//-----------------------------------------------------------------------------------------------------------------------------------------
// PRC 03 Cell loading
//-----------------------------------------------------------------------------------------------------------------------------------------
FOR nStationParameter := 20 TO 35
DO
  GVL_XTS.StationParameter[nStationParameter].rVelo               := 1000.0; //MAIN_APP.rDefaultVeloMin;
END_FOR
nStationParameter := 20;
GVL_XTS.StationParameter[nStationParameter].eType                 := E_STATION_TYPE.STATION_PROCESS;
GVL_XTS.StationParameter[nStationParameter].sText                 := 'PROCESS_INFEED_01';
GVL_XTS.StationParameter[nStationParameter].nConfiguredStopCount  :=       1;   // how many stops the mover has to make in this station

GVL_XTS.StationParameter[nStationParameter].rPosWait              :=    10000.0+80.0; // absolute modulo position
GVL_XTS.StationParameter[nStationParameter].rPosStop[1]           :=       0.0; // relative to rPosWait
GVL_XTS.StationParameter[nStationParameter].rReleaseDistance      :=    1120.0; // relative to Mover.ActPos

nStationParameter := 21;
GVL_XTS.StationParameter[nStationParameter].eType                 := E_STATION_TYPE.STATION_PROCESS;
GVL_XTS.StationParameter[nStationParameter].sText                 := 'PROCESS_INFEED_02';
GVL_XTS.StationParameter[nStationParameter].nConfiguredStopCount  :=       1;   // how many stops the mover has to make in this station

GVL_XTS.StationParameter[nStationParameter].rPosWait              :=    10000.0+160.0; // absolute modulo position
GVL_XTS.StationParameter[nStationParameter].rPosStop[1]           :=       0.0; // relative to rPosWait
GVL_XTS.StationParameter[nStationParameter].rReleaseDistance      :=    1040.0; // relative to Mover.ActPos

nStationParameter := 22;
GVL_XTS.StationParameter[nStationParameter].eType                 := E_STATION_TYPE.STATION_PROCESS;
GVL_XTS.StationParameter[nStationParameter].sText                 := 'PROCESS_INFEED_03';
GVL_XTS.StationParameter[nStationParameter].nConfiguredStopCount  :=       1;   // how many stops the mover has to make in this station

GVL_XTS.StationParameter[nStationParameter].rPosWait              :=    10000.0+240.0; // absolute modulo position
GVL_XTS.StationParameter[nStationParameter].rPosStop[1]           :=       0.0; // relative to rPosWait
GVL_XTS.StationParameter[nStationParameter].rReleaseDistance      :=     960.0; // relative to Mover.ActPos

nStationParameter := 23;
GVL_XTS.StationParameter[nStationParameter].eType                 := E_STATION_TYPE.STATION_PROCESS;
GVL_XTS.StationParameter[nStationParameter].sText                 := 'PROCESS_INFEED_04';
GVL_XTS.StationParameter[nStationParameter].nConfiguredStopCount  :=       1;   // how many stops the mover has to make in this station

GVL_XTS.StationParameter[nStationParameter].rPosWait              :=    10000.0+320.0; // absolute modulo position
GVL_XTS.StationParameter[nStationParameter].rPosStop[1]           :=       0.0; // relative to rPosWait
GVL_XTS.StationParameter[nStationParameter].rReleaseDistance      :=     880.0; // relative to Mover.ActPos

nStationParameter := 24;
GVL_XTS.StationParameter[nStationParameter].eType                 := E_STATION_TYPE.STATION_PROCESS;
GVL_XTS.StationParameter[nStationParameter].sText                 := 'PROCESS_INFEED_05';
GVL_XTS.StationParameter[nStationParameter].nConfiguredStopCount  :=       1;   // how many stops the mover has to make in this station

GVL_XTS.StationParameter[nStationParameter].rPosWait              :=    10000.0+400.0; // absolute modulo position
GVL_XTS.StationParameter[nStationParameter].rPosStop[1]           :=       0.0; // relative to rPosWait
GVL_XTS.StationParameter[nStationParameter].rReleaseDistance      :=     800.0; // relative to Mover.ActPos

nStationParameter := 25;
GVL_XTS.StationParameter[nStationParameter].eType                 := E_STATION_TYPE.STATION_PROCESS;
GVL_XTS.StationParameter[nStationParameter].sText                 := 'PROCESS_INFEED_06';
GVL_XTS.StationParameter[nStationParameter].nConfiguredStopCount  :=       1;   // how many stops the mover has to make in this station

GVL_XTS.StationParameter[nStationParameter].rPosWait              :=    10000.0+480.0; // absolute modulo position
GVL_XTS.StationParameter[nStationParameter].rPosStop[1]           :=       0.0; // relative to rPosWait
GVL_XTS.StationParameter[nStationParameter].rReleaseDistance      :=     720.0; // relative to Mover.ActPos

nStationParameter := 26;
GVL_XTS.StationParameter[nStationParameter].eType                 := E_STATION_TYPE.STATION_PROCESS;
GVL_XTS.StationParameter[nStationParameter].sText                 := 'PROCESS_INFEED_07';
GVL_XTS.StationParameter[nStationParameter].nConfiguredStopCount  :=       1;   // how many stops the mover has to make in this station

GVL_XTS.StationParameter[nStationParameter].rPosWait              :=    10000.0+560.0; // absolute modulo position
GVL_XTS.StationParameter[nStationParameter].rPosStop[1]           :=       0.0; // relative to rPosWait
GVL_XTS.StationParameter[nStationParameter].rReleaseDistance      :=     640.0; // relative to Mover.ActPos

nStationParameter := 27;
GVL_XTS.StationParameter[nStationParameter].eType                 := E_STATION_TYPE.STATION_PROCESS;
GVL_XTS.StationParameter[nStationParameter].sText                 := 'PROCESS_INFEED_08';
GVL_XTS.StationParameter[nStationParameter].nConfiguredStopCount  :=       1;   // how many stops the mover has to make in this station

GVL_XTS.StationParameter[nStationParameter].rPosWait              :=    10000.0+640.0; // absolute modulo position
GVL_XTS.StationParameter[nStationParameter].rPosStop[1]           :=       0.0; // relative to rPosWait
GVL_XTS.StationParameter[nStationParameter].rReleaseDistance      :=     560.0; // relative to Mover.ActPos

nStationParameter := 28;
GVL_XTS.StationParameter[nStationParameter].eType                 := E_STATION_TYPE.STATION_PROCESS;
GVL_XTS.StationParameter[nStationParameter].sText                 := 'PROCESS_INFEED_09';
GVL_XTS.StationParameter[nStationParameter].nConfiguredStopCount  :=       1;   // how many stops the mover has to make in this station

GVL_XTS.StationParameter[nStationParameter].rPosWait              :=    10000.0+720.0; // absolute modulo position
GVL_XTS.StationParameter[nStationParameter].rPosStop[1]           :=       0.0; // relative to rPosWait
GVL_XTS.StationParameter[nStationParameter].rReleaseDistance      :=     480.0; // relative to Mover.ActPos

nStationParameter := 29;
GVL_XTS.StationParameter[nStationParameter].eType                 := E_STATION_TYPE.STATION_PROCESS;
GVL_XTS.StationParameter[nStationParameter].sText                 := 'PROCESS_INFEED_10';
GVL_XTS.StationParameter[nStationParameter].nConfiguredStopCount  :=       1;   // how many stops the mover has to make in this station

GVL_XTS.StationParameter[nStationParameter].rPosWait              :=    10000.0+800.0; // absolute modulo position
GVL_XTS.StationParameter[nStationParameter].rPosStop[1]           :=       0.0; // relative to rPosWait
GVL_XTS.StationParameter[nStationParameter].rReleaseDistance      :=     400.0; // relative to Mover.ActPos

nStationParameter := 30;
GVL_XTS.StationParameter[nStationParameter].eType                 := E_STATION_TYPE.STATION_PROCESS;
GVL_XTS.StationParameter[nStationParameter].sText                 := 'PROCESS_INFEED_11';
GVL_XTS.StationParameter[nStationParameter].nConfiguredStopCount  :=       1;   // how many stops the mover has to make in this station

GVL_XTS.StationParameter[nStationParameter].rPosWait              :=    10000.0+880.0; // absolute modulo position
GVL_XTS.StationParameter[nStationParameter].rPosStop[1]           :=       0.0; // relative to rPosWait
GVL_XTS.StationParameter[nStationParameter].rReleaseDistance      :=     320.0; // relative to Mover.ActPos

nStationParameter := 31;
GVL_XTS.StationParameter[nStationParameter].eType                 := E_STATION_TYPE.STATION_PROCESS;
GVL_XTS.StationParameter[nStationParameter].sText                 := 'PROCESS_INFEED_12';
GVL_XTS.StationParameter[nStationParameter].nConfiguredStopCount  :=       1;   // how many stops the mover has to make in this station

GVL_XTS.StationParameter[nStationParameter].rPosWait              :=    10000.0+960.0; // absolute modulo position
GVL_XTS.StationParameter[nStationParameter].rPosStop[1]           :=       0.0; // relative to rPosWait
GVL_XTS.StationParameter[nStationParameter].rReleaseDistance      :=     240.0; // relative to Mover.ActPos

nStationParameter := 32;
GVL_XTS.StationParameter[nStationParameter].eType                 := E_STATION_TYPE.STATION_PROCESS;
GVL_XTS.StationParameter[nStationParameter].sText                 := 'PROCESS_INFEED_13';
GVL_XTS.StationParameter[nStationParameter].nConfiguredStopCount  :=       1;   // how many stops the mover has to make in this station

GVL_XTS.StationParameter[nStationParameter].rPosWait              :=    10000.0+1040.0; // absolute modulo position
GVL_XTS.StationParameter[nStationParameter].rPosStop[1]           :=       0.0; // relative to rPosWait
GVL_XTS.StationParameter[nStationParameter].rReleaseDistance      :=     160.0; // relative to Mover.ActPos

nStationParameter := 33;
GVL_XTS.StationParameter[nStationParameter].eType                 := E_STATION_TYPE.STATION_PROCESS;
GVL_XTS.StationParameter[nStationParameter].sText                 := 'PROCESS_INFEED_14';
GVL_XTS.StationParameter[nStationParameter].nConfiguredStopCount  :=       1;   // how many stops the mover has to make in this station

GVL_XTS.StationParameter[nStationParameter].rPosWait              :=    10000.0+1120.0; // absolute modulo position
GVL_XTS.StationParameter[nStationParameter].rPosStop[1]           :=       0.0; // relative to rPosWait
GVL_XTS.StationParameter[nStationParameter].rReleaseDistance      :=      80.0; // relative to Mover.ActPos

nStationParameter := 34;
GVL_XTS.StationParameter[nStationParameter].eType                 := E_STATION_TYPE.STATION_PROCESS;
GVL_XTS.StationParameter[nStationParameter].sText                 := 'PROCESS_INFEED_15';
GVL_XTS.StationParameter[nStationParameter].nConfiguredStopCount  :=       1;   // how many stops the mover has to make in this station

GVL_XTS.StationParameter[nStationParameter].rPosWait              :=    10000.0+1200.0; // absolute modulo position
GVL_XTS.StationParameter[nStationParameter].rPosStop[1]           :=       0.0; // relative to rPosWait
GVL_XTS.StationParameter[nStationParameter].rReleaseDistance      :=      25.0; // relative to Mover.ActPos

nStationParameter := 35;
GVL_XTS.StationParameter[nStationParameter].eType                 := E_STATION_TYPE.STATION_PROCESS;
GVL_XTS.StationParameter[nStationParameter].sText                 := 'PROCESS_INFEED_16';
GVL_XTS.StationParameter[nStationParameter].nConfiguredStopCount  :=       1;   // how many stops the mover has to make in this station

GVL_XTS.StationParameter[nStationParameter].rPosWait              :=    10000.0+1280.0; // absolute modulo position
GVL_XTS.StationParameter[nStationParameter].rPosStop[1]           :=       0.0; // relative to rPosWait
GVL_XTS.StationParameter[nStationParameter].rReleaseDistance      :=      -5.0; // relative to Mover.ActPos

//-----------------------------------------------------------------------------------------------------------------------------------------
// CONTINUOUS_CLEAN
//-----------------------------------------------------------------------------------------------------------------------------------------
nStationParameter := 37;
GVL_XTS.StationParameter[nStationParameter].eType                 := E_STATION_TYPE.STATION_PROCESS;
GVL_XTS.StationParameter[nStationParameter].sText                 := 'CONTINUOUS_CLEAN';
GVL_XTS.StationParameter[nStationParameter].nConfiguredStopCount  :=       1;   // how many stops the mover has to make in this station

GVL_XTS.StationParameter[nStationParameter].rPosWait              :=   12900.0; // absolute modulo position
GVL_XTS.StationParameter[nStationParameter].rPosStop[1]           :=       0.0; // relative to rPosWait
GVL_XTS.StationParameter[nStationParameter].rReleaseDistance      :=      -5.0; // relative to Mover.ActPos
GVL_XTS.StationParameter[nStationParameter].rVelo                 :=     250.0;
GVL_XTS.StationParameter[nStationParameter].rGap                  :=     110.0;

//-----------------------------------------------------------------------------------------------------------------------------------------
// CONTINUOUS_SCAN
//-----------------------------------------------------------------------------------------------------------------------------------------
nStationParameter := 38;
GVL_XTS.StationParameter[nStationParameter].eType                 := E_STATION_TYPE.STATION_PROCESS;
GVL_XTS.StationParameter[nStationParameter].sText                 := 'CONTINUOUS_SCAN';
GVL_XTS.StationParameter[nStationParameter].nConfiguredStopCount  :=       1;   // how many stops the mover has to make in this station

GVL_XTS.StationParameter[nStationParameter].rPosWait              :=   14000.0; // absolute modulo position
GVL_XTS.StationParameter[nStationParameter].rPosStop[1]           :=       0.0; // relative to rPosWait
GVL_XTS.StationParameter[nStationParameter].rReleaseDistance      :=      -5.0; // relative to Mover.ActPos
GVL_XTS.StationParameter[nStationParameter].rVelo                 :=     250.0;
GVL_XTS.StationParameter[nStationParameter].rGap                  :=     110.0;

//-----------------------------------------------------------------------------------------------------------------------------------------
// CONTINUOUS_CAM
//-----------------------------------------------------------------------------------------------------------------------------------------
nStationParameter := 39;
GVL_XTS.StationParameter[nStationParameter].eType                 := E_STATION_TYPE.STATION_PROCESS;
GVL_XTS.StationParameter[nStationParameter].sText                 := 'CONTINUOUS_CAM';
GVL_XTS.StationParameter[nStationParameter].nConfiguredStopCount  :=       1;   // how many stops the mover has to make in this station

GVL_XTS.StationParameter[nStationParameter].rPosWait              :=   14300.0; // absolute modulo position
GVL_XTS.StationParameter[nStationParameter].rPosStop[1]           :=       0.0; // relative to rPosWait
GVL_XTS.StationParameter[nStationParameter].rReleaseDistance      :=      -5.0; // relative to Mover.ActPos
GVL_XTS.StationParameter[nStationParameter].rVelo                 :=     250.0;
GVL_XTS.StationParameter[nStationParameter].rGap                  :=     109.0;

//-----------------------------------------------------------------------------------------------------------------------------------------
// DISTRIBUTOR_ASSEMBLY_01
//-----------------------------------------------------------------------------------------------------------------------------------------
nStationParameter := 40;
GVL_XTS.StationParameter[nStationParameter].eType                 := E_STATION_TYPE.STATION_PROCESS;
GVL_XTS.StationParameter[nStationParameter].sText                 := 'DISTRIBUTOR_ASSEMBLY_01';
GVL_XTS.StationParameter[nStationParameter].nConfiguredStopCount  :=       1;   // how many stops the mover has to make in this station

GVL_XTS.StationParameter[nStationParameter].rPosWait              :=   15250.0; // absolute modulo position
GVL_XTS.StationParameter[nStationParameter].rPosStop[1]           :=       0.0; // relative to rPosWait
GVL_XTS.StationParameter[nStationParameter].rReleaseDistance      :=      -5.0; // relative to Mover.ActPos
GVL_XTS.StationParameter[nStationParameter].rVelo                 :=    1500.0;
GVL_XTS.StationParameter[nStationParameter].rGap                  :=     109.0;

//-----------------------------------------------------------------------------------------------------------------------------------------
// PRC 05 Visual check film bottom
//-----------------------------------------------------------------------------------------------------------------------------------------
FOR nStationParameter := 41 TO 56
DO
  GVL_XTS.StationParameter[nStationParameter].rVelo               := MAIN_APP.rDefaultVeloMin;
END_FOR
nStationParameter := 41;
GVL_XTS.StationParameter[nStationParameter].eType                 := E_STATION_TYPE.STATION_PROCESS;
GVL_XTS.StationParameter[nStationParameter].sText                 := 'PROCESS_ASSEMBLY_01_01';
GVL_XTS.StationParameter[nStationParameter].nConfiguredStopCount  :=       1;   // how many stops the mover has to make in this station

GVL_XTS.StationParameter[nStationParameter].rPosWait              :=    15500.0+110.0; // absolute modulo position
GVL_XTS.StationParameter[nStationParameter].rPosStop[1]           :=       0.0; // relative to rPosWait
GVL_XTS.StationParameter[nStationParameter].rReleaseDistance      :=    1100.0; // relative to Mover.ActPos
GVL_XTS.StationParameter[nStationParameter].rGap                  :=     109.0;

nStationParameter := 42;
GVL_XTS.StationParameter[nStationParameter].eType                 := E_STATION_TYPE.STATION_PROCESS;
GVL_XTS.StationParameter[nStationParameter].sText                 := 'PROCESS_ASSEMBLY_01_02';
GVL_XTS.StationParameter[nStationParameter].nConfiguredStopCount  :=       1;   // how many stops the mover has to make in this station

GVL_XTS.StationParameter[nStationParameter].rPosWait              :=    15500.0+220.0; // absolute modulo position
GVL_XTS.StationParameter[nStationParameter].rPosStop[1]           :=       0.0; // relative to rPosWait
GVL_XTS.StationParameter[nStationParameter].rReleaseDistance      :=     990.0; // relative to Mover.ActPos
GVL_XTS.StationParameter[nStationParameter].rGap                  :=     109.0;

nStationParameter := 43;
GVL_XTS.StationParameter[nStationParameter].eType                 := E_STATION_TYPE.STATION_PROCESS;
GVL_XTS.StationParameter[nStationParameter].sText                 := 'PROCESS_ASSEMBLY_01_03';
GVL_XTS.StationParameter[nStationParameter].nConfiguredStopCount  :=       1;   // how many stops the mover has to make in this station

GVL_XTS.StationParameter[nStationParameter].rPosWait              :=    15500.0+330.0; // absolute modulo position
GVL_XTS.StationParameter[nStationParameter].rPosStop[1]           :=       0.0; // relative to rPosWait
GVL_XTS.StationParameter[nStationParameter].rReleaseDistance      :=     880.0; // relative to Mover.ActPos
GVL_XTS.StationParameter[nStationParameter].rGap                  :=     109.0;

nStationParameter := 44;
GVL_XTS.StationParameter[nStationParameter].eType                 := E_STATION_TYPE.STATION_PROCESS;
GVL_XTS.StationParameter[nStationParameter].sText                 := 'PROCESS_ASSEMBLY_01_04';
GVL_XTS.StationParameter[nStationParameter].nConfiguredStopCount  :=       1;   // how many stops the mover has to make in this station

GVL_XTS.StationParameter[nStationParameter].rPosWait              :=    15500.0+440.0; // absolute modulo position
GVL_XTS.StationParameter[nStationParameter].rPosStop[1]           :=       0.0; // relative to rPosWait
GVL_XTS.StationParameter[nStationParameter].rReleaseDistance      :=     770.0; // relative to Mover.ActPos
GVL_XTS.StationParameter[nStationParameter].rGap                  :=     109.0;

nStationParameter := 45;
GVL_XTS.StationParameter[nStationParameter].eType                 := E_STATION_TYPE.STATION_PROCESS;
GVL_XTS.StationParameter[nStationParameter].sText                 := 'PROCESS_ASSEMBLY_01_05';
GVL_XTS.StationParameter[nStationParameter].nConfiguredStopCount  :=       1;   // how many stops the mover has to make in this station

GVL_XTS.StationParameter[nStationParameter].rPosWait              :=    15500.0+550.0; // absolute modulo position
GVL_XTS.StationParameter[nStationParameter].rPosStop[1]           :=       0.0; // relative to rPosWait
GVL_XTS.StationParameter[nStationParameter].rReleaseDistance      :=     660.0; // relative to Mover.ActPos
GVL_XTS.StationParameter[nStationParameter].rGap                  :=     109.0;

nStationParameter := 46;
GVL_XTS.StationParameter[nStationParameter].eType                 := E_STATION_TYPE.STATION_PROCESS;
GVL_XTS.StationParameter[nStationParameter].sText                 := 'PROCESS_ASSEMBLY_01_06';
GVL_XTS.StationParameter[nStationParameter].nConfiguredStopCount  :=       1;   // how many stops the mover has to make in this station

GVL_XTS.StationParameter[nStationParameter].rPosWait              :=    15500.0+660.0; // absolute modulo position
GVL_XTS.StationParameter[nStationParameter].rPosStop[1]           :=       0.0; // relative to rPosWait
GVL_XTS.StationParameter[nStationParameter].rReleaseDistance      :=     550.0; // relative to Mover.ActPos
GVL_XTS.StationParameter[nStationParameter].rGap                  :=     109.0;

nStationParameter := 47;
GVL_XTS.StationParameter[nStationParameter].eType                 := E_STATION_TYPE.STATION_PROCESS;
GVL_XTS.StationParameter[nStationParameter].sText                 := 'PROCESS_ASSEMBLY_01_07';
GVL_XTS.StationParameter[nStationParameter].nConfiguredStopCount  :=       1;   // how many stops the mover has to make in this station

GVL_XTS.StationParameter[nStationParameter].rPosWait              :=    15500.0+770.0; // absolute modulo position
GVL_XTS.StationParameter[nStationParameter].rPosStop[1]           :=       0.0; // relative to rPosWait
GVL_XTS.StationParameter[nStationParameter].rReleaseDistance      :=     440.0; // relative to Mover.ActPos
GVL_XTS.StationParameter[nStationParameter].rGap                  :=     109.0;

nStationParameter := 48;
GVL_XTS.StationParameter[nStationParameter].eType                 := E_STATION_TYPE.STATION_PROCESS;
GVL_XTS.StationParameter[nStationParameter].sText                 := 'PROCESS_ASSEMBLY_01_08';
GVL_XTS.StationParameter[nStationParameter].nConfiguredStopCount  :=       1;   // how many stops the mover has to make in this station

GVL_XTS.StationParameter[nStationParameter].rPosWait              :=    15500.0+880.0; // absolute modulo position
GVL_XTS.StationParameter[nStationParameter].rPosStop[1]           :=       0.0; // relative to rPosWait
GVL_XTS.StationParameter[nStationParameter].rReleaseDistance      :=     330.0; // relative to Mover.ActPos
GVL_XTS.StationParameter[nStationParameter].rGap                  :=     109.0;

nStationParameter := 49;
GVL_XTS.StationParameter[nStationParameter].eType                 := E_STATION_TYPE.STATION_PROCESS;
GVL_XTS.StationParameter[nStationParameter].sText                 := 'PROCESS_ASSEMBLY_01_09';
GVL_XTS.StationParameter[nStationParameter].nConfiguredStopCount  :=       1;   // how many stops the mover has to make in this station

GVL_XTS.StationParameter[nStationParameter].rPosWait              :=    15500.0+990.0; // absolute modulo position
GVL_XTS.StationParameter[nStationParameter].rPosStop[1]           :=       0.0; // relative to rPosWait
GVL_XTS.StationParameter[nStationParameter].rReleaseDistance      :=     220.0; // relative to Mover.ActPos
GVL_XTS.StationParameter[nStationParameter].rGap                  :=     109.0;

nStationParameter := 50;
GVL_XTS.StationParameter[nStationParameter].eType                 := E_STATION_TYPE.STATION_PROCESS;
GVL_XTS.StationParameter[nStationParameter].sText                 := 'PROCESS_ASSEMBLY_01_10';
GVL_XTS.StationParameter[nStationParameter].nConfiguredStopCount  :=       1;   // how many stops the mover has to make in this station
GVL_XTS.StationParameter[nStationParameter].rGap                  :=     110.0;

GVL_XTS.StationParameter[nStationParameter].rPosWait              :=    15500.0+1100.0; // absolute modulo position
GVL_XTS.StationParameter[nStationParameter].rPosStop[1]           :=       0.0; // relative to rPosWait
GVL_XTS.StationParameter[nStationParameter].rReleaseDistance      :=     110.0; // relative to Mover.ActPos
GVL_XTS.StationParameter[nStationParameter].rGap                  :=     109.0;

nStationParameter := 51;
GVL_XTS.StationParameter[nStationParameter].eType                 := E_STATION_TYPE.STATION_PROCESS;
GVL_XTS.StationParameter[nStationParameter].sText                 := 'PROCESS_ASSEMBLY_01_11';
GVL_XTS.StationParameter[nStationParameter].nConfiguredStopCount  :=       1;   // how many stops the mover has to make in this station

GVL_XTS.StationParameter[nStationParameter].rPosWait              :=    15500.0+1210.0; // absolute modulo position
GVL_XTS.StationParameter[nStationParameter].rPosStop[1]           :=       0.0; // relative to rPosWait
GVL_XTS.StationParameter[nStationParameter].rReleaseDistance      :=     25.0; // relative to Mover.ActPos
GVL_XTS.StationParameter[nStationParameter].rGap                  :=     109.0;

nStationParameter := 52;
GVL_XTS.StationParameter[nStationParameter].eType                 := E_STATION_TYPE.STATION_PROCESS;
GVL_XTS.StationParameter[nStationParameter].sText                 := 'PROCESS_ASSEMBLY_01_12';
GVL_XTS.StationParameter[nStationParameter].nConfiguredStopCount  :=       1;   // how many stops the mover has to make in this station

GVL_XTS.StationParameter[nStationParameter].rPosWait              :=    15500.0+1320.0; // absolute modulo position
GVL_XTS.StationParameter[nStationParameter].rPosStop[1]           :=       0.0; // relative to rPosWait
GVL_XTS.StationParameter[nStationParameter].rReleaseDistance      :=     330.0; // relative to Mover.ActPos
GVL_XTS.StationParameter[nStationParameter].rGap                  :=     109.0;

nStationParameter := 53;
GVL_XTS.StationParameter[nStationParameter].eType                 := E_STATION_TYPE.STATION_PROCESS;
GVL_XTS.StationParameter[nStationParameter].sText                 := 'PROCESS_ASSEMBLY_01_13';
GVL_XTS.StationParameter[nStationParameter].nConfiguredStopCount  :=       1;   // how many stops the mover has to make in this station

GVL_XTS.StationParameter[nStationParameter].rPosWait              :=    15500.0+1430.0; // absolute modulo position
GVL_XTS.StationParameter[nStationParameter].rPosStop[1]           :=       0.0; // relative to rPosWait
GVL_XTS.StationParameter[nStationParameter].rReleaseDistance      :=     220.0; // relative to Mover.ActPos
GVL_XTS.StationParameter[nStationParameter].rGap                  :=     109.0;

nStationParameter := 54;
GVL_XTS.StationParameter[nStationParameter].eType                 := E_STATION_TYPE.STATION_PROCESS;
GVL_XTS.StationParameter[nStationParameter].sText                 := 'PROCESS_ASSEMBLY_01_14';
GVL_XTS.StationParameter[nStationParameter].nConfiguredStopCount  :=       1;   // how many stops the mover has to make in this station

GVL_XTS.StationParameter[nStationParameter].rPosWait              :=    15500.0+1540.0; // absolute modulo position
GVL_XTS.StationParameter[nStationParameter].rPosStop[1]           :=       0.0; // relative to rPosWait
GVL_XTS.StationParameter[nStationParameter].rReleaseDistance      :=     110.0; // relative to Mover.ActPos
GVL_XTS.StationParameter[nStationParameter].rGap                  :=     109.0;

nStationParameter := 55;
GVL_XTS.StationParameter[nStationParameter].eType                 := E_STATION_TYPE.STATION_PROCESS;
GVL_XTS.StationParameter[nStationParameter].sText                 := 'PROCESS_ASSEMBLY_01_15';
GVL_XTS.StationParameter[nStationParameter].nConfiguredStopCount  :=       1;   // how many stops the mover has to make in this station

GVL_XTS.StationParameter[nStationParameter].rPosWait              :=    15500.0+1650.0; // absolute modulo position
GVL_XTS.StationParameter[nStationParameter].rPosStop[1]           :=       0.0; // relative to rPosWait
GVL_XTS.StationParameter[nStationParameter].rReleaseDistance      :=      25.0; // relative to Mover.ActPos
GVL_XTS.StationParameter[nStationParameter].rGap                  :=     109.0;

nStationParameter := 56;
GVL_XTS.StationParameter[nStationParameter].eType                 := E_STATION_TYPE.STATION_PROCESS;
GVL_XTS.StationParameter[nStationParameter].sText                 := 'PROCESS_ASSEMBLY_01_16';
GVL_XTS.StationParameter[nStationParameter].nConfiguredStopCount  :=       1;   // how many stops the mover has to make in this station

GVL_XTS.StationParameter[nStationParameter].rPosWait              :=    15500.0+1740.0; // absolute modulo position
GVL_XTS.StationParameter[nStationParameter].rPosStop[1]           :=       0.0; // relative to rPosWait
GVL_XTS.StationParameter[nStationParameter].rReleaseDistance      :=      -5.0; // relative to Mover.ActPos
GVL_XTS.StationParameter[nStationParameter].rGap                  :=     109.0;
//-----------------------------------------------------------------------------------------------------------------------------------------
// DISTRIBUTOR_ASSEMBLY_02
//-----------------------------------------------------------------------------------------------------------------------------------------
nStationParameter := 57;
GVL_XTS.StationParameter[nStationParameter].eType                 := E_STATION_TYPE.STATION_PROCESS;
GVL_XTS.StationParameter[nStationParameter].sText                 := 'DISTRIBUTOR_ASSEMBLY_02';
GVL_XTS.StationParameter[nStationParameter].nConfiguredStopCount  :=       1;   // how many stops the mover has to make in this station

GVL_XTS.StationParameter[nStationParameter].rPosWait              :=   18000.0; // absolute modulo position
GVL_XTS.StationParameter[nStationParameter].rPosStop[1]           :=       0.0; // relative to rPosWait
GVL_XTS.StationParameter[nStationParameter].rReleaseDistance      :=      -5.0; // relative to Mover.ActPos
GVL_XTS.StationParameter[nStationParameter].rVelo                 := MAIN_APP.rDefaultVeloMin;

//-----------------------------------------------------------------------------------------------------------------------------------------
// PROCESS_ASSEMBLY_02
//-----------------------------------------------------------------------------------------------------------------------------------------
FOR nStationParameter := 58 TO 69
DO
   GVL_XTS.StationParameter[nStationParameter].rVelo               := MAIN_APP.rDefaultVeloMin;
END_FOR
nStationParameter := 58;
GVL_XTS.StationParameter[nStationParameter].eType                 := E_STATION_TYPE.STATION_PROCESS;
GVL_XTS.StationParameter[nStationParameter].sText                 := 'PROCESS_ASSEMBLY_02_01';
GVL_XTS.StationParameter[nStationParameter].nConfiguredStopCount  :=       1;   // how many stops the mover has to make in this station

GVL_XTS.StationParameter[nStationParameter].rPosWait              :=    19500.0+80.0; // absolute modulo position
GVL_XTS.StationParameter[nStationParameter].rPosStop[1]           :=       0.0; // relative to rPosWait
GVL_XTS.StationParameter[nStationParameter].rReleaseDistance      :=     480.0; // relative to Mover.ActPos

nStationParameter := 59;
GVL_XTS.StationParameter[nStationParameter].eType                 := E_STATION_TYPE.STATION_PROCESS;
GVL_XTS.StationParameter[nStationParameter].sText                 := 'PROCESS_ASSEMBLY_02_02';
GVL_XTS.StationParameter[nStationParameter].nConfiguredStopCount  :=       1;   // how many stops the mover has to make in this station

GVL_XTS.StationParameter[nStationParameter].rPosWait              :=    19500.0+160.0; // absolute modulo position
GVL_XTS.StationParameter[nStationParameter].rPosStop[1]           :=       0.0; // relative to rPosWait
GVL_XTS.StationParameter[nStationParameter].rReleaseDistance      :=     400.0; // relative to Mover.ActPos

nStationParameter := 60;
GVL_XTS.StationParameter[nStationParameter].eType                 := E_STATION_TYPE.STATION_PROCESS;
GVL_XTS.StationParameter[nStationParameter].sText                 := 'PROCESS_ASSEMBLY_02_03';
GVL_XTS.StationParameter[nStationParameter].nConfiguredStopCount  :=       1;   // how many stops the mover has to make in this station

GVL_XTS.StationParameter[nStationParameter].rPosWait              :=    19500.0+240.0; // absolute modulo position
GVL_XTS.StationParameter[nStationParameter].rPosStop[1]           :=       0.0; // relative to rPosWait
GVL_XTS.StationParameter[nStationParameter].rReleaseDistance      :=     320.0; // relative to Mover.ActPos

nStationParameter := 61;
GVL_XTS.StationParameter[nStationParameter].eType                 := E_STATION_TYPE.STATION_PROCESS;
GVL_XTS.StationParameter[nStationParameter].sText                 := 'PROCESS_ASSEMBLY_02_04';
GVL_XTS.StationParameter[nStationParameter].nConfiguredStopCount  :=       1;   // how many stops the mover has to make in this station

GVL_XTS.StationParameter[nStationParameter].rPosWait              :=    19500.0+320.0; // absolute modulo position
GVL_XTS.StationParameter[nStationParameter].rPosStop[1]           :=       0.0; // relative to rPosWait
GVL_XTS.StationParameter[nStationParameter].rReleaseDistance      :=     240.0; // relative to Mover.ActPos

nStationParameter := 62;
GVL_XTS.StationParameter[nStationParameter].eType                 := E_STATION_TYPE.STATION_PROCESS;
GVL_XTS.StationParameter[nStationParameter].sText                 := 'PROCESS_ASSEMBLY_02_05';
GVL_XTS.StationParameter[nStationParameter].nConfiguredStopCount  :=       1;   // how many stops the mover has to make in this station

GVL_XTS.StationParameter[nStationParameter].rPosWait              :=    19500.0+400.0; // absolute modulo position
GVL_XTS.StationParameter[nStationParameter].rPosStop[1]           :=       0.0; // relative to rPosWait
GVL_XTS.StationParameter[nStationParameter].rReleaseDistance      :=      160.0; // relative to Mover.ActPos

nStationParameter := 63;
GVL_XTS.StationParameter[nStationParameter].eType                 := E_STATION_TYPE.STATION_PROCESS;
GVL_XTS.StationParameter[nStationParameter].sText                 := 'PROCESS_ASSEMBLY_02_06';
GVL_XTS.StationParameter[nStationParameter].nConfiguredStopCount  :=       1;   // how many stops the mover has to make in this station

GVL_XTS.StationParameter[nStationParameter].rPosWait              :=    19500.0+480.0; // absolute modulo position
GVL_XTS.StationParameter[nStationParameter].rPosStop[1]           :=       0.0; // relative to rPosWait
GVL_XTS.StationParameter[nStationParameter].rReleaseDistance      :=      80.0; // relative to Mover.ActPos

nStationParameter := 64;
GVL_XTS.StationParameter[nStationParameter].eType                 := E_STATION_TYPE.STATION_PROCESS;
GVL_XTS.StationParameter[nStationParameter].sText                 := 'PROCESS_ASSEMBLY_02_07';
GVL_XTS.StationParameter[nStationParameter].nConfiguredStopCount  :=       1;   // how many stops the mover has to make in this station

GVL_XTS.StationParameter[nStationParameter].rPosWait              :=    19500.0+560.0; // absolute modulo position
GVL_XTS.StationParameter[nStationParameter].rPosStop[1]           :=       0.0; // relative to rPosWait
GVL_XTS.StationParameter[nStationParameter].rReleaseDistance      :=      25.0; // relative to Mover.ActPos

nStationParameter := 65;
GVL_XTS.StationParameter[nStationParameter].eType                 := E_STATION_TYPE.STATION_PROCESS;
GVL_XTS.StationParameter[nStationParameter].sText                 := 'PROCESS_ASSEMBLY_02_08';
GVL_XTS.StationParameter[nStationParameter].nConfiguredStopCount  :=       1;   // how many stops the mover has to make in this station

GVL_XTS.StationParameter[nStationParameter].rPosWait              :=    19500.0+640.0; // absolute modulo position
GVL_XTS.StationParameter[nStationParameter].rPosStop[1]           :=       0.0; // relative to rPosWait
GVL_XTS.StationParameter[nStationParameter].rReleaseDistance      :=     -5.0; // relative to Mover.ActPos

nStationParameter := 66;
GVL_XTS.StationParameter[nStationParameter].eType                 := E_STATION_TYPE.STATION_PROCESS;
GVL_XTS.StationParameter[nStationParameter].sText                 := 'PROCESS_ASSEMBLY_02_09';
GVL_XTS.StationParameter[nStationParameter].nConfiguredStopCount  :=       1;   // how many stops the mover has to make in this station

GVL_XTS.StationParameter[nStationParameter].rPosWait              :=    19500.0+720.0; // absolute modulo position
GVL_XTS.StationParameter[nStationParameter].rPosStop[1]           :=       0.0; // relative to rPosWait
GVL_XTS.StationParameter[nStationParameter].rReleaseDistance      :=     240.0; // relative to Mover.ActPos

nStationParameter := 67;
GVL_XTS.StationParameter[nStationParameter].eType                 := E_STATION_TYPE.STATION_PROCESS;
GVL_XTS.StationParameter[nStationParameter].sText                 := 'PROCESS_ASSEMBLY_02_10';
GVL_XTS.StationParameter[nStationParameter].nConfiguredStopCount  :=       1;   // how many stops the mover has to make in this station

GVL_XTS.StationParameter[nStationParameter].rPosWait              :=    19500.0+800.0; // absolute modulo position
GVL_XTS.StationParameter[nStationParameter].rPosStop[1]           :=       0.0; // relative to rPosWait
GVL_XTS.StationParameter[nStationParameter].rReleaseDistance      :=     160.0; // relative to Mover.ActPos

nStationParameter := 68;
GVL_XTS.StationParameter[nStationParameter].eType                 := E_STATION_TYPE.STATION_PROCESS;
GVL_XTS.StationParameter[nStationParameter].sText                 := 'PROCESS_ASSEMBLY_02_11';
GVL_XTS.StationParameter[nStationParameter].nConfiguredStopCount  :=       1;   // how many stops the mover has to make in this station

GVL_XTS.StationParameter[nStationParameter].rPosWait              :=    19500.0+880.0; // absolute modulo position
GVL_XTS.StationParameter[nStationParameter].rPosStop[1]           :=       0.0; // relative to rPosWait
GVL_XTS.StationParameter[nStationParameter].rReleaseDistance      :=      80.0; // relative to Mover.ActPos

nStationParameter := 69;
GVL_XTS.StationParameter[nStationParameter].eType                 := E_STATION_TYPE.STATION_PROCESS;
GVL_XTS.StationParameter[nStationParameter].sText                 := 'PROCESS_ASSEMBLY_02_12';
GVL_XTS.StationParameter[nStationParameter].nConfiguredStopCount  :=       1;   // how many stops the mover has to make in this station

GVL_XTS.StationParameter[nStationParameter].rPosWait              :=    19500.0+960.0; // absolute modulo position
GVL_XTS.StationParameter[nStationParameter].rPosStop[1]           :=       0.0; // relative to rPosWait
GVL_XTS.StationParameter[nStationParameter].rReleaseDistance      :=      25.0; // relative to Mover.ActPos

//-----------------------------------------------------------------------------------------------------------------------------------------
// DISTRIBUTOR_ASSEMBLY_TEST
//-----------------------------------------------------------------------------------------------------------------------------------------
nStationParameter := 70;
GVL_XTS.StationParameter[nStationParameter].eType                 := E_STATION_TYPE.STATION_PROCESS;
GVL_XTS.StationParameter[nStationParameter].sText                 := 'DISTRIBUTOR_ASSEMBLY_TEST';
GVL_XTS.StationParameter[nStationParameter].nConfiguredStopCount  :=       1;   // how many stops the mover has to make in this station

GVL_XTS.StationParameter[nStationParameter].rPosWait              :=   21000.0; // absolute modulo position
GVL_XTS.StationParameter[nStationParameter].rPosStop[1]           :=       0.0; // relative to rPosWait
GVL_XTS.StationParameter[nStationParameter].rReleaseDistance      :=      -5.0; // relative to Mover.ActPos


//-----------------------------------------------------------------------------------------------------------------------------------------
// PROCESS_ASSEMBLY_TEST
//-----------------------------------------------------------------------------------------------------------------------------------------
FOR nStationParameter := 71 TO 86
DO
   GVL_XTS.StationParameter[nStationParameter].rVelo               := 1000.0;//MAIN_APP.rDefaultVeloMin;
END_FOR
nStationParameter := 71;
GVL_XTS.StationParameter[nStationParameter].eType                 := E_STATION_TYPE.STATION_PROCESS;
GVL_XTS.StationParameter[nStationParameter].sText                 := 'PROCESS_ASSEMBLY_TEST_01';
GVL_XTS.StationParameter[nStationParameter].nConfiguredStopCount  :=       1;   // how many stops the mover has to make in this station

GVL_XTS.StationParameter[nStationParameter].rPosWait              :=    21500.0+80.0; // absolute modulo position
GVL_XTS.StationParameter[nStationParameter].rPosStop[1]           :=       0.0; // relative to rPosWait
GVL_XTS.StationParameter[nStationParameter].rReleaseDistance      :=     800.0; // relative to Mover.ActPos

nStationParameter := 72;
GVL_XTS.StationParameter[nStationParameter].eType                 := E_STATION_TYPE.STATION_PROCESS;
GVL_XTS.StationParameter[nStationParameter].sText                 := 'PROCESS_ASSEMBLY_TEST_02';
GVL_XTS.StationParameter[nStationParameter].nConfiguredStopCount  :=       1;   // how many stops the mover has to make in this station

GVL_XTS.StationParameter[nStationParameter].rPosWait              :=    21500.0+160.0; // absolute modulo position
GVL_XTS.StationParameter[nStationParameter].rPosStop[1]           :=       0.0; // relative to rPosWait
GVL_XTS.StationParameter[nStationParameter].rReleaseDistance      :=     720.0; // relative to Mover.ActPos

nStationParameter := 73;
GVL_XTS.StationParameter[nStationParameter].eType                 := E_STATION_TYPE.STATION_PROCESS;
GVL_XTS.StationParameter[nStationParameter].sText                 := 'PROCESS_ASSEMBLY_TEST_03';
GVL_XTS.StationParameter[nStationParameter].nConfiguredStopCount  :=       1;   // how many stops the mover has to make in this station

GVL_XTS.StationParameter[nStationParameter].rPosWait              :=    21500.0+240.0; // absolute modulo position
GVL_XTS.StationParameter[nStationParameter].rPosStop[1]           :=       0.0; // relative to rPosWait
GVL_XTS.StationParameter[nStationParameter].rReleaseDistance      :=    640.0; // relative to Mover.ActPos

nStationParameter := 74;
GVL_XTS.StationParameter[nStationParameter].eType                 := E_STATION_TYPE.STATION_PROCESS;
GVL_XTS.StationParameter[nStationParameter].sText                 := 'PROCESS_ASSEMBLY_TEST_04';
GVL_XTS.StationParameter[nStationParameter].nConfiguredStopCount  :=       1;   // how many stops the mover has to make in this station

GVL_XTS.StationParameter[nStationParameter].rPosWait              :=    21500.0+320.0; // absolute modulo position
GVL_XTS.StationParameter[nStationParameter].rPosStop[1]           :=       0.0; // relative to rPosWait
GVL_XTS.StationParameter[nStationParameter].rReleaseDistance      :=     560.0; // relative to Mover.ActPos

nStationParameter := 75;
GVL_XTS.StationParameter[nStationParameter].eType                 := E_STATION_TYPE.STATION_PROCESS;
GVL_XTS.StationParameter[nStationParameter].sText                 := 'PROCESS_ASSEMBLY_TEST_05';
GVL_XTS.StationParameter[nStationParameter].nConfiguredStopCount  :=       1;   // how many stops the mover has to make in this station

GVL_XTS.StationParameter[nStationParameter].rPosWait              :=    21500.0+400.0; // absolute modulo position
GVL_XTS.StationParameter[nStationParameter].rPosStop[1]           :=       0.0; // relative to rPosWait
GVL_XTS.StationParameter[nStationParameter].rReleaseDistance      :=     480.0; // relative to Mover.ActPos

nStationParameter := 76;
GVL_XTS.StationParameter[nStationParameter].eType                 := E_STATION_TYPE.STATION_PROCESS;
GVL_XTS.StationParameter[nStationParameter].sText                 := 'PROCESS_ASSEMBLY_TEST_06';
GVL_XTS.StationParameter[nStationParameter].nConfiguredStopCount  :=       1;   // how many stops the mover has to make in this station

GVL_XTS.StationParameter[nStationParameter].rPosWait              :=    21500.0+480.0; // absolute modulo position
GVL_XTS.StationParameter[nStationParameter].rPosStop[1]           :=       0.0; // relative to rPosWait
GVL_XTS.StationParameter[nStationParameter].rReleaseDistance      :=     400.0; // relative to Mover.ActPos

nStationParameter := 77;
GVL_XTS.StationParameter[nStationParameter].eType                 := E_STATION_TYPE.STATION_PROCESS;
GVL_XTS.StationParameter[nStationParameter].sText                 := 'PROCESS_ASSEMBLY_TEST_07';
GVL_XTS.StationParameter[nStationParameter].nConfiguredStopCount  :=       1;   // how many stops the mover has to make in this station

GVL_XTS.StationParameter[nStationParameter].rPosWait              :=    21500.0+560.0; // absolute modulo position
GVL_XTS.StationParameter[nStationParameter].rPosStop[1]           :=       0.0; // relative to rPosWait
GVL_XTS.StationParameter[nStationParameter].rReleaseDistance      :=     320.0; // relative to Mover.ActPos

nStationParameter := 78;
GVL_XTS.StationParameter[nStationParameter].eType                 := E_STATION_TYPE.STATION_PROCESS;
GVL_XTS.StationParameter[nStationParameter].sText                 := 'PROCESS_ASSEMBLY_TEST_08';
GVL_XTS.StationParameter[nStationParameter].nConfiguredStopCount  :=       1;   // how many stops the mover has to make in this station

GVL_XTS.StationParameter[nStationParameter].rPosWait              :=    21500.0+640.0; // absolute modulo position
GVL_XTS.StationParameter[nStationParameter].rPosStop[1]           :=       0.0; // relative to rPosWait
GVL_XTS.StationParameter[nStationParameter].rReleaseDistance      :=     240.0; // relative to Mover.ActPos

nStationParameter := 79;
GVL_XTS.StationParameter[nStationParameter].eType                 := E_STATION_TYPE.STATION_PROCESS;
GVL_XTS.StationParameter[nStationParameter].sText                 := 'PROCESS_ASSEMBLY_TEST_09';
GVL_XTS.StationParameter[nStationParameter].nConfiguredStopCount  :=       1;   // how many stops the mover has to make in this station

GVL_XTS.StationParameter[nStationParameter].rPosWait              :=    21500.0+720.0; // absolute modulo position
GVL_XTS.StationParameter[nStationParameter].rPosStop[1]           :=       0.0; // relative to rPosWait
GVL_XTS.StationParameter[nStationParameter].rReleaseDistance      :=     160.0; // relative to Mover.ActPos

nStationParameter := 80;
GVL_XTS.StationParameter[nStationParameter].eType                 := E_STATION_TYPE.STATION_PROCESS;
GVL_XTS.StationParameter[nStationParameter].sText                 := 'PROCESS_ASSEMBLY_TEST_10';
GVL_XTS.StationParameter[nStationParameter].nConfiguredStopCount  :=       1;   // how many stops the mover has to make in this station

GVL_XTS.StationParameter[nStationParameter].rPosWait              :=    21500.0+800.0; // absolute modulo position
GVL_XTS.StationParameter[nStationParameter].rPosStop[1]           :=       0.0; // relative to rPosWait
GVL_XTS.StationParameter[nStationParameter].rReleaseDistance      :=      80.0; // relative to Mover.ActPos

nStationParameter := 81;
GVL_XTS.StationParameter[nStationParameter].eType                 := E_STATION_TYPE.STATION_PROCESS;
GVL_XTS.StationParameter[nStationParameter].sText                 := 'PROCESS_ASSEMBLY_TEST_11';
GVL_XTS.StationParameter[nStationParameter].nConfiguredStopCount  :=       1;   // how many stops the mover has to make in this station

GVL_XTS.StationParameter[nStationParameter].rPosWait              :=    21500.0+880.0; // absolute modulo position
GVL_XTS.StationParameter[nStationParameter].rPosStop[1]           :=       0.0; // relative to rPosWait
GVL_XTS.StationParameter[nStationParameter].rReleaseDistance      :=      25.0; // relative to Mover.ActPos

nStationParameter := 82;
GVL_XTS.StationParameter[nStationParameter].eType                 := E_STATION_TYPE.STATION_PROCESS;
GVL_XTS.StationParameter[nStationParameter].sText                 := 'PROCESS_ASSEMBLY_TEST_12';
GVL_XTS.StationParameter[nStationParameter].nConfiguredStopCount  :=       1;   // how many stops the mover has to make in this station

GVL_XTS.StationParameter[nStationParameter].rPosWait              :=    21500.0+960.0; // absolute modulo position
GVL_XTS.StationParameter[nStationParameter].rPosStop[1]           :=       0.0; // relative to rPosWait
GVL_XTS.StationParameter[nStationParameter].rReleaseDistance      :=     -5.0; // relative to Mover.ActPos

nStationParameter := 83;
GVL_XTS.StationParameter[nStationParameter].eType                 := E_STATION_TYPE.STATION_PROCESS;
GVL_XTS.StationParameter[nStationParameter].sText                 := 'PROCESS_ASSEMBLY_TEST_13';
GVL_XTS.StationParameter[nStationParameter].nConfiguredStopCount  :=       1;   // how many stops the mover has to make in this station

GVL_XTS.StationParameter[nStationParameter].rPosWait              :=    21500.0+1040.0; // absolute modulo position
GVL_XTS.StationParameter[nStationParameter].rPosStop[1]           :=       0.0; // relative to rPosWait
GVL_XTS.StationParameter[nStationParameter].rReleaseDistance      :=     240.0; // relative to Mover.ActPos

nStationParameter := 84;
GVL_XTS.StationParameter[nStationParameter].eType                 := E_STATION_TYPE.STATION_PROCESS;
GVL_XTS.StationParameter[nStationParameter].sText                 := 'PRC_08_1_14_HV_TEST';
GVL_XTS.StationParameter[nStationParameter].nConfiguredStopCount  :=       1;   // how many stops the mover has to make in this station

GVL_XTS.StationParameter[nStationParameter].rPosWait              :=    21500.0+1120.0; // absolute modulo position
GVL_XTS.StationParameter[nStationParameter].rPosStop[1]           :=       0.0; // relative to rPosWait
GVL_XTS.StationParameter[nStationParameter].rReleaseDistance      :=     160.0; // relative to Mover.ActPos

nStationParameter := 85;
GVL_XTS.StationParameter[nStationParameter].eType                 := E_STATION_TYPE.STATION_PROCESS;
GVL_XTS.StationParameter[nStationParameter].sText                 := 'PRC_08_1_15_HV_TEST';
GVL_XTS.StationParameter[nStationParameter].nConfiguredStopCount  :=       1;   // how many stops the mover has to make in this station

GVL_XTS.StationParameter[nStationParameter].rPosWait              :=    21500.0+1200.0; // absolute modulo position
GVL_XTS.StationParameter[nStationParameter].rPosStop[1]           :=       0.0; // relative to rPosWait
GVL_XTS.StationParameter[nStationParameter].rReleaseDistance      :=      80.0; // relative to Mover.ActPos

nStationParameter := 86;
GVL_XTS.StationParameter[nStationParameter].eType                 := E_STATION_TYPE.STATION_PROCESS;
GVL_XTS.StationParameter[nStationParameter].sText                 := 'PRC_08_1_16_HV_TEST';
GVL_XTS.StationParameter[nStationParameter].nConfiguredStopCount  :=       1;   // how many stops the mover has to make in this station

GVL_XTS.StationParameter[nStationParameter].rPosWait              :=    21500.0+1280.0; // absolute modulo position
GVL_XTS.StationParameter[nStationParameter].rPosStop[1]           :=       0.0; // relative to rPosWait
GVL_XTS.StationParameter[nStationParameter].rReleaseDistance      :=      25.0; // relative to Mover.ActPos

//-----------------------------------------------------------------------------------------------------------------------------------------
// NOK handling
//-----------------------------------------------------------------------------------------------------------------------------------------
FOR nStationParameter := 91 TO 91
DO
  GVL_XTS.StationParameter[nStationParameter].rVelo               := 750.0;//MAIN_APP.rDefaultVeloMin;
END_FOR
nStationParameter := 91;
GVL_XTS.StationParameter[nStationParameter].eType                 := E_STATION_TYPE.STATION_PROCESS;
GVL_XTS.StationParameter[nStationParameter].sText                 := 'PRC_09_NOK';
GVL_XTS.StationParameter[nStationParameter].nConfiguredStopCount  :=       1;   // how many stops the mover has to make in this station

GVL_XTS.StationParameter[nStationParameter].rPosWait              :=   23250.0; // absolute modulo position
GVL_XTS.StationParameter[nStationParameter].rPosStop[1]           :=       0.0; // relative to rPosWait
GVL_XTS.StationParameter[nStationParameter].rReleaseDistance      :=      -5.0; // relative to Mover.ActPos

//-----------------------------------------------------------------------------------------------------------------------------------------
// PRC 09 CELL CLEANING 
//-----------------------------------------------------------------------------------------------------------------------------------------
FOR nStationParameter := 95 TO 95
DO
  GVL_XTS.StationParameter[nStationParameter].rVelo               := MAIN_APP.rDefaultVeloMin;
END_FOR
nStationParameter := 95;
GVL_XTS.StationParameter[nStationParameter].eType                 := E_STATION_TYPE.STATION_PROCESS;
GVL_XTS.StationParameter[nStationParameter].sText                 := 'PRC_09_CELL_CLEANING';
GVL_XTS.StationParameter[nStationParameter].nConfiguredStopCount  :=       1;   // how many stops the mover has to make in this station

GVL_XTS.StationParameter[nStationParameter].rPosWait              :=   24000.0+80.0; // absolute modulo position
GVL_XTS.StationParameter[nStationParameter].rPosStop[1]           :=       0.0; // relative to rPosWait
GVL_XTS.StationParameter[nStationParameter].rReleaseDistance      :=      -5.0; // relative to Mover.ActPos
GVL_XTS.StationParameter[nStationParameter].rVelo                 :=     750.0;
GVL_XTS.StationParameter[nStationParameter].rGap                  :=      78.0;

//-----------------------------------------------------------------------------------------------------------------------------------------
// DISTRIBUTOR - cell unloading
//-----------------------------------------------------------------------------------------------------------------------------------------
nStationParameter := 119;
GVL_XTS.StationParameter[nStationParameter].eType                 := E_STATION_TYPE.STATION_PROCESS;
GVL_XTS.StationParameter[nStationParameter].sText                 := 'DIST_12_CELL_UNLOAD';
GVL_XTS.StationParameter[nStationParameter].nConfiguredStopCount  :=       1;   // how many stops the mover has to make in this station

GVL_XTS.StationParameter[nStationParameter].rPosWait              :=   26000.0; // absolute modulo position
GVL_XTS.StationParameter[nStationParameter].rPosStop[1]           :=       0.0; // relative to rPosWait
GVL_XTS.StationParameter[nStationParameter].rReleaseDistance      :=      -5.0; // relative to Mover.ActPos
GVL_XTS.StationParameter[nStationParameter].rVelo                 :=    1000.0;//MAIN_APP.rDefaultVeloMin;


//-----------------------------------------------------------------------------------------------------------------------------------------
// PROCESS_OUTFEED
//-----------------------------------------------------------------------------------------------------------------------------------------
FOR nStationParameter := 120 TO 133
DO
  GVL_XTS.StationParameter[nStationParameter].rVelo               := 1000.0;//MAIN_APP.rDefaultVeloMin;
END_FOR
nStationParameter := 120;
GVL_XTS.StationParameter[nStationParameter].eType                 := E_STATION_TYPE.STATION_PROCESS;
GVL_XTS.StationParameter[nStationParameter].sText                 := 'PROCESS_OUTFEED_01';
GVL_XTS.StationParameter[nStationParameter].nConfiguredStopCount  :=       1;   // how many stops the mover has to make in this station

GVL_XTS.StationParameter[nStationParameter].rPosWait              :=   26250.0; // absolute modulo position
GVL_XTS.StationParameter[nStationParameter].rPosStop[1]           :=      80.0; // relative to rPosWait
GVL_XTS.StationParameter[nStationParameter].rReleaseDistance      :=     960.0; // relative to Mover.ActPos

nStationParameter := 121;
GVL_XTS.StationParameter[nStationParameter].eType                 := E_STATION_TYPE.STATION_PROCESS;
GVL_XTS.StationParameter[nStationParameter].sText                 := 'PROCESS_OUTFEED_02';
GVL_XTS.StationParameter[nStationParameter].nConfiguredStopCount  :=       1;   // how many stops the mover has to make in this station

GVL_XTS.StationParameter[nStationParameter].rPosWait              :=   26250.0; // absolute modulo position
GVL_XTS.StationParameter[nStationParameter].rPosStop[1]           :=     160.0; // relative to rPosWait
GVL_XTS.StationParameter[nStationParameter].rReleaseDistance      :=     880.0; // relative to Mover.ActPos

nStationParameter := 122;
GVL_XTS.StationParameter[nStationParameter].eType                 := E_STATION_TYPE.STATION_PROCESS;
GVL_XTS.StationParameter[nStationParameter].sText                 := 'PROCESS_OUTFEED_03';
GVL_XTS.StationParameter[nStationParameter].nConfiguredStopCount  :=       1;   // how many stops the mover has to make in this station

GVL_XTS.StationParameter[nStationParameter].rPosWait              :=   26250.0; // absolute modulo position
GVL_XTS.StationParameter[nStationParameter].rPosStop[1]           :=     240.0; // relative to rPosWait
GVL_XTS.StationParameter[nStationParameter].rReleaseDistance      :=     800.0; // relative to Mover.ActPos

nStationParameter := 123;
GVL_XTS.StationParameter[nStationParameter].eType                 := E_STATION_TYPE.STATION_PROCESS;
GVL_XTS.StationParameter[nStationParameter].sText                 := 'PROCESS_OUTFEED_04';
GVL_XTS.StationParameter[nStationParameter].nConfiguredStopCount  :=       1;   // how many stops the mover has to make in this station

GVL_XTS.StationParameter[nStationParameter].rPosWait              :=   26250.0; // absolute modulo position
GVL_XTS.StationParameter[nStationParameter].rPosStop[1]           :=     320.0; // relative to rPosWait
GVL_XTS.StationParameter[nStationParameter].rReleaseDistance      :=     720.0; // relative to Mover.ActPos

nStationParameter := 124;
GVL_XTS.StationParameter[nStationParameter].eType                 := E_STATION_TYPE.STATION_PROCESS;
GVL_XTS.StationParameter[nStationParameter].sText                 := 'PROCESS_OUTFEED_05';
GVL_XTS.StationParameter[nStationParameter].nConfiguredStopCount  :=       1;   // how many stops the mover has to make in this station

GVL_XTS.StationParameter[nStationParameter].rPosWait              :=   26250.0; // absolute modulo position
GVL_XTS.StationParameter[nStationParameter].rPosStop[1]           :=     400.0; // relative to rPosWait
GVL_XTS.StationParameter[nStationParameter].rReleaseDistance      :=     640.0; // relative to Mover.ActPos

nStationParameter := 125;
GVL_XTS.StationParameter[nStationParameter].eType                 := E_STATION_TYPE.STATION_PROCESS;
GVL_XTS.StationParameter[nStationParameter].sText                 := 'PROCESS_OUTFEED_06';
GVL_XTS.StationParameter[nStationParameter].nConfiguredStopCount  :=       1;   // how many stops the mover has to make in this station

GVL_XTS.StationParameter[nStationParameter].rPosWait              :=   26250.0; // absolute modulo position
GVL_XTS.StationParameter[nStationParameter].rPosStop[1]           :=     480.0; // relative to rPosWait
GVL_XTS.StationParameter[nStationParameter].rReleaseDistance      :=     560.0; // relative to Mover.ActPos

nStationParameter := 126;
GVL_XTS.StationParameter[nStationParameter].eType                 := E_STATION_TYPE.STATION_PROCESS;
GVL_XTS.StationParameter[nStationParameter].sText                 := 'PROCESS_OUTFEED_07';
GVL_XTS.StationParameter[nStationParameter].nConfiguredStopCount  :=       1;   // how many stops the mover has to make in this station

GVL_XTS.StationParameter[nStationParameter].rPosWait              :=   26250.0; // absolute modulo position
GVL_XTS.StationParameter[nStationParameter].rPosStop[1]           :=     560.0; // relative to rPosWait
GVL_XTS.StationParameter[nStationParameter].rReleaseDistance      :=     480.0; // relative to Mover.ActPos

nStationParameter := 127;
GVL_XTS.StationParameter[nStationParameter].eType                 := E_STATION_TYPE.STATION_PROCESS;
GVL_XTS.StationParameter[nStationParameter].sText                 := 'PROCESS_OUTFEED_08';
GVL_XTS.StationParameter[nStationParameter].nConfiguredStopCount  :=       1;   // how many stops the mover has to make in this station

GVL_XTS.StationParameter[nStationParameter].rPosWait              :=   26250.0; // absolute modulo position
GVL_XTS.StationParameter[nStationParameter].rPosStop[1]           :=     640.0; // relative to rPosWait
GVL_XTS.StationParameter[nStationParameter].rReleaseDistance      :=     400.0; // relative to Mover.ActPos

nStationParameter := 128;
GVL_XTS.StationParameter[nStationParameter].eType                 := E_STATION_TYPE.STATION_PROCESS;
GVL_XTS.StationParameter[nStationParameter].sText                 := 'PROCESS_OUTFEED_09';
GVL_XTS.StationParameter[nStationParameter].nConfiguredStopCount  :=       1;   // how many stops the mover has to make in this station

GVL_XTS.StationParameter[nStationParameter].rPosWait              :=   26250.0; // absolute modulo position
GVL_XTS.StationParameter[nStationParameter].rPosStop[1]           :=     720.0; // relative to rPosWait
GVL_XTS.StationParameter[nStationParameter].rReleaseDistance      :=     320.0; // relative to Mover.ActPos

nStationParameter := 129;
GVL_XTS.StationParameter[nStationParameter].eType                 := E_STATION_TYPE.STATION_PROCESS;
GVL_XTS.StationParameter[nStationParameter].sText                 := 'PROCESS_OUTFEED_10';
GVL_XTS.StationParameter[nStationParameter].nConfiguredStopCount  :=       1;   // how many stops the mover has to make in this station

GVL_XTS.StationParameter[nStationParameter].rPosWait              :=   26250.0; // absolute modulo position
GVL_XTS.StationParameter[nStationParameter].rPosStop[1]           :=     800.0; // relative to rPosWait
GVL_XTS.StationParameter[nStationParameter].rReleaseDistance      :=     240.0; // relative to Mover.ActPos

nStationParameter := 130;
GVL_XTS.StationParameter[nStationParameter].eType                 := E_STATION_TYPE.STATION_PROCESS;
GVL_XTS.StationParameter[nStationParameter].sText                 := 'PROCESS_OUTFEED_11';
GVL_XTS.StationParameter[nStationParameter].nConfiguredStopCount  :=       1;   // how many stops the mover has to make in this station

GVL_XTS.StationParameter[nStationParameter].rPosWait              :=   26250.0; // absolute modulo position
GVL_XTS.StationParameter[nStationParameter].rPosStop[1]           :=     880.0; // relative to rPosWait
GVL_XTS.StationParameter[nStationParameter].rReleaseDistance      :=     160.0; // relative to Mover.ActPos

nStationParameter := 131;
GVL_XTS.StationParameter[nStationParameter].eType                 := E_STATION_TYPE.STATION_PROCESS;
GVL_XTS.StationParameter[nStationParameter].sText                 := 'PROCESS_OUTFEED_12';
GVL_XTS.StationParameter[nStationParameter].nConfiguredStopCount  :=       1;   // how many stops the mover has to make in this station

GVL_XTS.StationParameter[nStationParameter].rPosWait              :=   26250.0; // absolute modulo position
GVL_XTS.StationParameter[nStationParameter].rPosStop[1]           :=     960.0; // relative to rPosWait
GVL_XTS.StationParameter[nStationParameter].rReleaseDistance      :=     80.0; // relative to Mover.ActPos

nStationParameter := 132;
GVL_XTS.StationParameter[nStationParameter].eType                 := E_STATION_TYPE.STATION_PROCESS;
GVL_XTS.StationParameter[nStationParameter].sText                 := 'PROCESS_OUTFEED_13';
GVL_XTS.StationParameter[nStationParameter].nConfiguredStopCount  :=       1;   // how many stops the mover has to make in this station

GVL_XTS.StationParameter[nStationParameter].rPosWait              :=   26250.0; // absolute modulo position
GVL_XTS.StationParameter[nStationParameter].rPosStop[1]           :=    1040.0; // relative to rPosWait
GVL_XTS.StationParameter[nStationParameter].rReleaseDistance      :=      25.0; // relative to Mover.ActPos

nStationParameter := 133;
GVL_XTS.StationParameter[nStationParameter].eType                 := E_STATION_TYPE.STATION_PROCESS;
GVL_XTS.StationParameter[nStationParameter].sText                 := 'PROCESS_OUTFEED_14';
GVL_XTS.StationParameter[nStationParameter].nConfiguredStopCount  :=       1;   // how many stops the mover has to make in this station

GVL_XTS.StationParameter[nStationParameter].rPosWait              :=   26250.0; // absolute modulo position
GVL_XTS.StationParameter[nStationParameter].rPosStop[1]           :=    1120.0; // relative to rPosWait
GVL_XTS.StationParameter[nStationParameter].rReleaseDistance      :=      -5.0; // relative to Mover.ActPos

//-----------------------------------------------------------------------------------------------------------------------------------------
//  DISTRIBUTOR
//-----------------------------------------------------------------------------------------------------------------------------------------
nStationParameter := 140;
GVL_XTS.StationParameter[nStationParameter].eType                 := E_STATION_TYPE.STATION_PROCESS;
GVL_XTS.StationParameter[nStationParameter].sText                 := 'DISTRIBUTOR_WPC_CLEAN';
GVL_XTS.StationParameter[nStationParameter].nConfiguredStopCount  :=      1;   // how many stops the mover has to make in this station

GVL_XTS.StationParameter[nStationParameter].rPosWait              :=   1000.0; // absolute modulo position
GVL_XTS.StationParameter[nStationParameter].rPosStop[1]           :=      0.0; // relative to rPosWait
GVL_XTS.StationParameter[nStationParameter].rReleaseDistance      :=     -5.0; // relative to Mover.ActPos

GVL_XTS.StationParameter[nStationParameter].rGap                  :=     78.0;
GVL_XTS.StationParameter[nStationParameter].rVelo                 :=   2500.0;
GVL_XTS.StationParameter[nStationParameter].rAccDec               :=  17500.0;
GVL_XTS.StationParameter[nStationParameter].rJerk                 :=  300000.0;

//-----------------------------------------------------------------------------------------------------------------------------------------
//  PRC 14 wpc clean
//-----------------------------------------------------------------------------------------------------------------------------------------
nStationParameter := 141;
GVL_XTS.StationParameter[nStationParameter].eType                 := E_STATION_TYPE.STATION_PROCESS;
GVL_XTS.StationParameter[nStationParameter].sText                 := 'CONTINUOUS_WPC_CLEAN';
GVL_XTS.StationParameter[nStationParameter].nConfiguredStopCount  :=      1;   // how many stops the mover has to make in this station

GVL_XTS.StationParameter[nStationParameter].rPosWait              :=   4000.0; // absolute modulo position
GVL_XTS.StationParameter[nStationParameter].rPosStop[1]           :=      0.0; // relative to rPosWait
GVL_XTS.StationParameter[nStationParameter].rReleaseDistance      :=      -5.0; // relative to Mover.ActPos
GVL_XTS.StationParameter[nStationParameter].rVelo                 :=     500.0;
GVL_XTS.StationParameter[nStationParameter].rGap                  :=      78.0;
GVL_XTS.StationParameter[nStationParameter].rJerk                 :=  300000.0;

//-----------------------------------------------------------------------------------------------------------------------------------------
//  DISTRIBUTOR
//-----------------------------------------------------------------------------------------------------------------------------------------
nStationParameter := 142;
GVL_XTS.StationParameter[nStationParameter].eType                 := E_STATION_TYPE.STATION_PROCESS;
GVL_XTS.StationParameter[nStationParameter].sText                 := 'DISTRIBUTOR_INFEED';
GVL_XTS.StationParameter[nStationParameter].nConfiguredStopCount  :=      1;   // how many stops the mover has to make in this station

GVL_XTS.StationParameter[nStationParameter].rPosWait              :=   5500.0; // absolute modulo position
GVL_XTS.StationParameter[nStationParameter].rPosStop[1]           :=      0.0; // relative to rPosWait
GVL_XTS.StationParameter[nStationParameter].rReleaseDistance      :=     -5.0; // relative to Mover.ActPos

GVL_XTS.StationParameter[nStationParameter].rGap                  :=     78.0;
GVL_XTS.StationParameter[nStationParameter].rVelo                 :=   2000.0;

//-----------------------------------------------------------------------------------------------------------------------------------------
//-----------------------------------------------------------------------------------------------------------------------------------------
// EOF
//-----------------------------------------------------------------------------------------------------------------------------------------
//-----------------------------------------------------------------------------------------------------------------------------------------

END_FUNCTION

// ---- APPLICATION/MAIN_APPLICATION.TcVIS
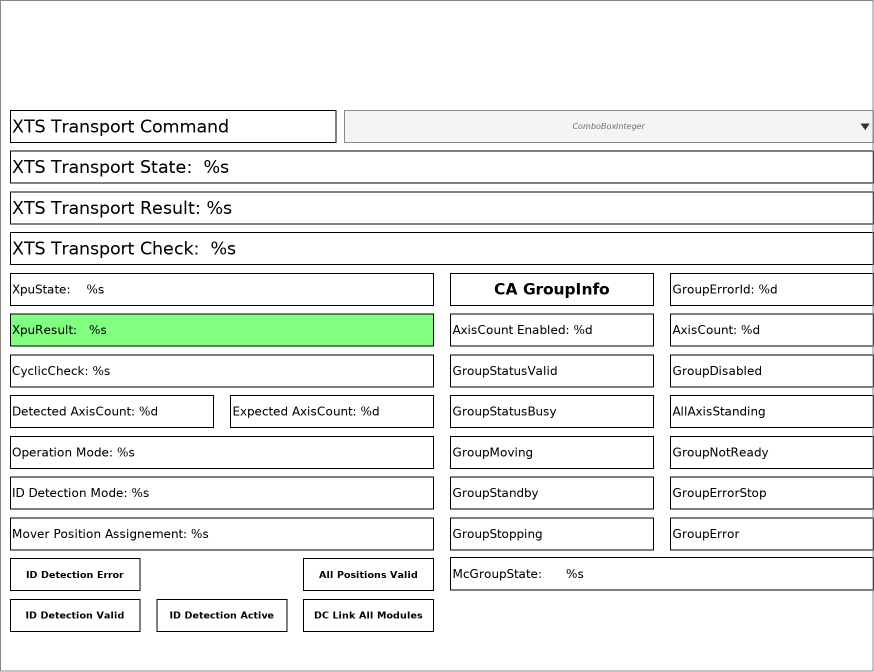
VISUALIZATION MAIN_APPLICATION  // 874x672
    Frame (10,110 864x562)
        shows TRANSPORT_VISU(Data := GVL_APPLICATION.VisuPoolData)
END_VISUALIZATION

// ---- APPLICATION/_Visualization/MOVER_VISU.TcVIS
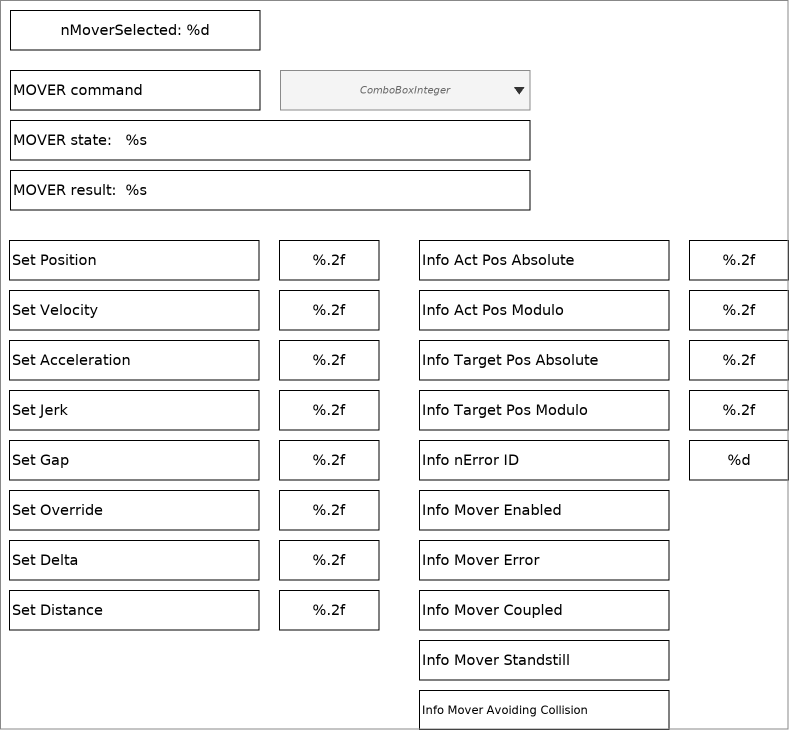
VISUALIZATION MOVER_VISU  // 789x730
    Rectangle (10,10 250x40), "nMoverSelected: %d", text variable: VISU_POOL.nMoverSelected
        OnMouseClick: write the text variable via VisuDialogs.Numpad, min 1, max MAX_MOVER, title 'Selected Mover'
    Rectangle (10,120 520x40), "MOVER state: %s", text variable: GVL_APPLICATION.VisuPoolData.sMoverState
    Rectangle (10,70 250x40), "MOVER command"
    ComboBoxInteger (280,70 250x40), variable: GVL_XTS.MoverCtrl[VISU_POOL.nMoverSelected].Cmd, text list: 'TL_E_CTRL_MOVER'
    Rectangle (10,170 520x40), "MOVER result: %s", text variable: GVL_APPLICATION.VisuPoolData.sMoverResult
    Rectangle (9,240 250x40), "Set Position"
    Rectangle (9,290 250x40), "Set Velocity"
    Rectangle (9,340 250x40), "Set Acceleration"
    Rectangle (9,390 250x40), "Set Jerk"
    Rectangle (9,440 250x40), "Set Gap"
    Rectangle (9,490 250x40), "Set Override"
    Rectangle (9,540 250x40), "Set Delta"
    Rectangle (9,590 250x40), "Set Distance"
    Rectangle (279,240 100x40), "%.2f", text variable: GVL_XTS.MoveData[VISU_POOL.nMoverSelected].rPos
        OnMouseClick: write the text variable via Default
    Rectangle (279,290 100x40), "%.2f", text variable: GVL_XTS.MoveData[VISU_POOL.nMoverSelected].rVelo
        OnMouseClick: write the text variable via Default
    Rectangle (279,340 100x40), "%.2f", text variable: GVL_XTS.MoveData[VISU_POOL.nMoverSelected].rAcc
        OnMouseClick: write the text variable via Default
    Rectangle (279,390 100x40), "%.2f", text variable: GVL_XTS.MoveData[VISU_POOL.nMoverSelected].rJerk
        OnMouseClick: write the text variable via Default
    Rectangle (279,440 100x40), "%.2f", text variable: GVL_XTS.MoveData[VISU_POOL.nMoverSelected].rGap
        OnMouseClick: write the text variable via Default
    Rectangle (279,490 100x40), "%.2f", text variable: GVL_XTS.MoveData[VISU_POOL.nMoverSelected].rOverride
        OnMouseClick: write the text variable via Default
    Rectangle (279,540 100x40), "%.2f", text variable: GVL_XTS.MoveData[VISU_POOL.nMoverSelected].rDelta
        OnMouseClick: write the text variable via Default
    Rectangle (279,590 100x40), "%.2f", text variable: GVL_XTS.MoveData[VISU_POOL.nMoverSelected].rDistance
        OnMouseClick: write the text variable via Default
    Rectangle (419,240 250x40), "Info Act Pos Absolute"
    Rectangle (419,290 250x40), "Info Act Pos Modulo"
    Rectangle (419,340 250x40), "Info Target Pos Absolute"
    Rectangle (419,390 250x40), "Info Target Pos Modulo"
    Rectangle (419,440 250x40), "Info nError ID"
    Rectangle (689,240 100x40), "%.2f", text variable: GVL_XTS.MoverInfo[VISU_POOL.nMoverSelected].rAbsActPos
    Rectangle (689,290 100x40), "%.2f", text variable: GVL_XTS.MoverInfo[VISU_POOL.nMoverSelected].rModuloActPos
    Rectangle (689,340 100x40), "%.2f", text variable: GVL_XTS.MoverInfo[VISU_POOL.nMoverSelected].rAbsTargetPos
    Rectangle (689,390 100x40), "%.2f", text variable: GVL_XTS.MoverInfo[VISU_POOL.nMoverSelected].rModuloTargetPos
    Rectangle (689,440 100x40), "%d", text variable: GVL_XTS.MoverInfo[VISU_POOL.nMoverSelected].nErrorId
    Rectangle (419,490 250x40), "Info Mover Enabled", colour toggle: GVL_XTS.MoverInfo[MAIN.nMoverSelected].bMoverEnabled
    Rectangle (419,540 250x40), "Info Mover Error", colour toggle: GVL_XTS.MoverInfo[MAIN.nMoverSelected].bMoverError
    Rectangle (419,590 250x40), "Info Mover Coupled", colour toggle: GVL_XTS.MoverInfo[MAIN.nMoverSelected].bMoverCoupled
    Rectangle (419,640 250x40), "Info Mover Standstill", colour toggle: GVL_XTS.MoverInfo[MAIN.nMoverSelected].bMoverStandstill
    Rectangle (419,690 250x40), "Info Mover Avoiding Collision", colour toggle: GVL_XTS.MoverInfo[MAIN.nMoverSelected].bMoverAvoidingCollision
END_VISUALIZATION

// ---- APPLICATION/_Visualization/SELECTOR_VISU.TcVIS
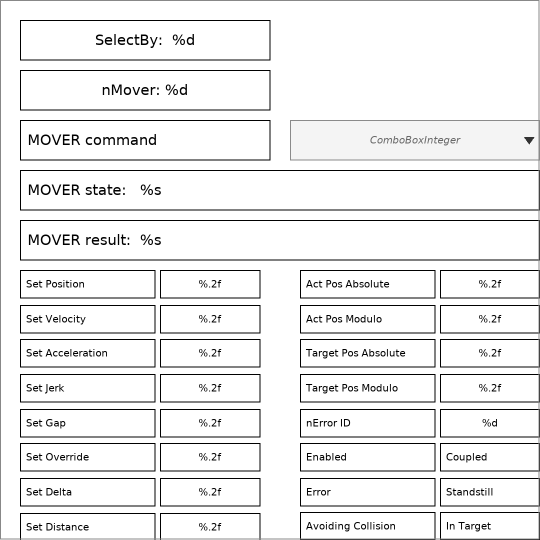
VISUALIZATION SELECTOR_VISU  // 540x540
    Frame (10,10 530x530)
        shows T_MOVER_SELECTOR(Control := GVL_XTS.MoverSelectorCtrl, State := GVL_XTS.MoverSelectorState, sState := GVL_APPLICATION.VisuPoolData.sSelectorState, sResult := GVL_APPLICATION.VisuPoolData.sSelectorResult)
END_VISUALIZATION

// ---- APPLICATION/_Visualization/STATION_VISU.TcVIS
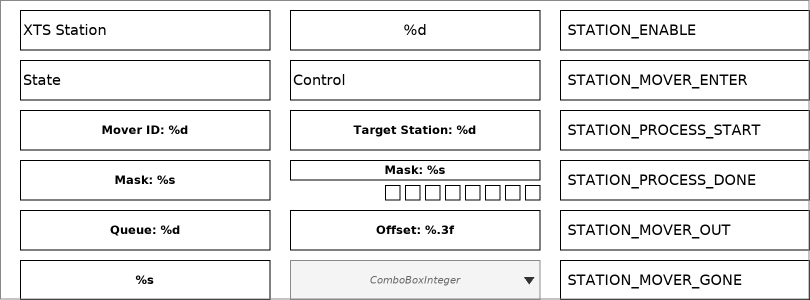
VISUALIZATION STATION_VISU  // 810x300
    Rectangle (20,10 250x40), "XTS Station"
    Rectangle (290,10 250x40), "%d", text variable: VISU_POOL.nStationSelected
        OnMouseClick: write the text variable via VisuDialogs.Numpad, min 1, max MAX_STATION, title 'Selected Station'
    Rectangle (20,60 250x40), "State"
    Rectangle (290,60 250x40), "Control"
    Rectangle (20,210 250x40), "Queue: %d", text variable: GVL_XTS.StationState[VISU_POOL.nStationSelected].nQueue
    Rectangle (20,110 250x40), "Mover ID: %d", text variable: GVL_XTS.StationState[VISU_POOL.nStationSelected].nMoverId
    Rectangle (20,160 250x40), "Mask: %s", text variable: GVL_APPLICATION.VisuPoolData.sStationStateMask
    Rectangle (20,260 250x40), "%s", text variable: GVL_APPLICATION.VisuPoolData.sStationState
    ComboBoxInteger (290,260 250x40), variable: GVL_XTS.StationCtrl[VISU_POOL.nStationSelected].eCmd, text list: 'TL_E_CTRL_STATION'
    Rectangle (290,210 250x40), "Offset: %.3f", text variable: GVL_XTS.StationCtrl[VISU_POOL.nStationSelected].rOffset
    Rectangle (290,110 250x40), "Target Station: %d", text variable: GVL_XTS.StationCtrl[VISU_POOL.nStationSelected].nTargetStation
        OnMouseClick: write the text variable via VisuDialogs.Numpad, min 1, max MAX_STATION, title 'Target Station'
    Rectangle (290,160 250x20), "Mask: %s", text variable: GVL_APPLICATION.VisuPoolData.sStationCtrlMask
    Rectangle (525,185 15x15)
        toggle GVL_XTS.StationCtrl[VISU_POOL.nStationSelected].nMask.0
    Rectangle (505,185 15x15)
        toggle GVL_XTS.StationCtrl[VISU_POOL.nStationSelected].nMask.1
    Rectangle (485,185 15x15)
        toggle GVL_XTS.StationCtrl[VISU_POOL.nStationSelected].nMask.2
    Rectangle (465,185 15x15)
        toggle GVL_XTS.StationCtrl[VISU_POOL.nStationSelected].nMask.3
    Rectangle (445,185 15x15)
        toggle GVL_XTS.StationCtrl[VISU_POOL.nStationSelected].nMask.4
    Rectangle (425,185 15x15)
        toggle GVL_XTS.StationCtrl[VISU_POOL.nStationSelected].nMask.5
    Rectangle (405,185 15x15)
        toggle GVL_XTS.StationCtrl[VISU_POOL.nStationSelected].nMask.6
    Rectangle (385,185 15x15)
        toggle GVL_XTS.StationCtrl[VISU_POOL.nStationSelected].nMask.7
    Rectangle (560,10 250x40), "STATION_ENABLE", colour toggle: GVL_APPLICATION.VisuPoolData.bStationEnable
        OnMouseClick: execute { GVL_XTS.StationCtrl[VISU_POOL.nMoverSelected].Cmd := E_STATION_CTRL.STATION_ENABLE; }
    Rectangle (560,60 250x40), "STATION_MOVER_ENTER", colour toggle: GVL_APPLICATION.VisuPoolData.bStationEnter
        OnMouseClick: execute { GVL_XTS.StationCtrl[VISU_POOL.nMoverSelected].Cmd := E_STATION_CTRL.STATION_MOVER_ENTER; }
    Rectangle (560,110 250x40), "STATION_PROCESS_START", colour toggle: GVL_APPLICATION.VisuPoolData.bStationStart
        OnMouseClick: execute { GVL_XTS.StationCtrl[VISU_POOL.nMoverSelected].Cmd := E_STATION_CTRL.STATION_PROCESS_START; }
    Rectangle (560,160 250x40), "STATION_PROCESS_DONE", colour toggle: GVL_APPLICATION.VisuPoolData.bStationDone
        OnMouseClick: execute { GVL_XTS.StationCtrl[VISU_POOL.nMoverSelected].Cmd := E_STATION_CTRL.STATION_PROCESS_DONE; }
    Rectangle (560,210 250x40), "STATION_MOVER_OUT", colour toggle: GVL_APPLICATION.VisuPoolData.bStationOut
        OnMouseClick: execute { GVL_XTS.StationCtrl[VISU_POOL.nMoverSelected].Cmd := E_STATION_CTRL.STATION_MOVER_OUT; }
    Rectangle (560,260 250x40), "STATION_MOVER_GONE", colour toggle: GVL_APPLICATION.VisuPoolData.bStationGone
        OnMouseClick: execute { GVL_XTS.StationCtrl[VISU_POOL.nMoverSelected].Cmd := E_STATION_CTRL.STATION_MOVER_GONE; }
END_VISUALIZATION

// ---- APPLICATION/_Visualization/TRANSPORT_VISU.TcVIS
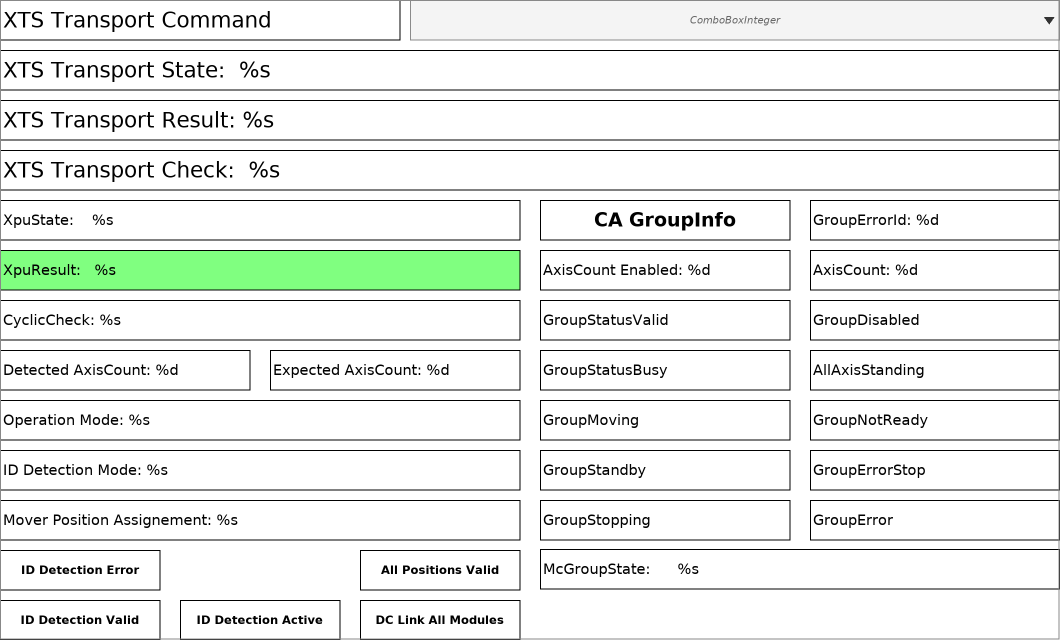
VISUALIZATION TRANSPORT_VISU  // 1060x640
VAR_IN_OUT
	Data    : ST_VISU_POOL;
END_VAR
    Rectangle (0,0 400x40), "XTS Transport Command"
    ComboBoxInteger (410,0 650x40), variable: GVL_XTS.XtsTransportCtrl.Cmd, text list: 'TL_E_CTRL_TRANSPORT'
    Rectangle (0,50 1060x40), "XTS Transport State: %s", text variable: Data.sTransportState
    Rectangle (0,100 1060x40), "XTS Transport Result: %s", text variable: Data.sTransportResult
    Rectangle (0,150 1060x40), "XTS Transport Check: %s", text variable: Data.sTransportCheck
    Frame (0,200 520x440)
        shows XPU_VISU(stXpuState := GVL_XTS.XtsTransportState.XpuState, stXpuInfo := GVL_XTS.XtsTransportState.XpuInfo, stXpuStrings := Data.stXpuStrings)
    Frame (540,200 520x390)
        shows GROUP_VISU(stGroupInfo := GVL_XTS.XtsTransportState.GroupInfo, sGroupState := Data.sCaGroupState)
END_VISUALIZATION

// ---- GlobalTextList.TcGTLO
TEXTLIST GlobalTextList
  230 = ' %d'
  30 = ' Act Pos Absolute'
  518 = ' Act Pos Modulo'
  493 = ' Avoiding Collision'
  587 = ' Coupled'
  690 = ' Enabled'
  968 = ' Error'
  733 = ' In Target'
  144 = ' MOVER command'
  271 = ' MOVER result:  %s'
  268 = ' MOVER state:   %s'
  484 = ' nError ID'
  912 = ' Set Acceleration'
  819 = ' Set Delta'
  464 = ' Set Distance'
  1025 = ' Set Gap'
  363 = ' Set Jerk'
  376 = ' Set Override'
  1069 = ' Set Position'
  859 = ' Set Velocity'
  123 = ' Standstill'
  17 = ' STATION_ENABLE'
  34 = ' STATION_MOVER_ENTER'
  452 = ' STATION_MOVER_GONE'
  75 = ' STATION_MOVER_OUT'
  598 = ' STATION_PROCESS_DONE'
  750 = ' STATION_PROCESS_START'
  727 = ' Target Pos Absolute'
  397 = ' Target Pos Modulo'
  294 = '%.2f'
  191 = '%d'
  836 = '%s'
  704 = 'All Positions Valid'
  562 = 'AllAxisStanding'
  878 = 'AxisCount Enabled: %d'
  162 = 'AxisCount: %d'
  516 = 'CA GroupInfo'
  929 = 'Control'
  707 = 'CyclicCheck: %s'
  660 = 'DC Link All Modules'
  843 = 'Detected AxisCount: %d'
  772 = 'Expected AxisCount: %d'
  48 = 'GroupDisabled'
  915 = 'GroupError'
  495 = 'GroupErrorId: %d'
  975 = 'GroupErrorStop'
  300 = 'GroupMoving'
  807 = 'GroupNotReady'
  438 = 'GroupStandby'
  226 = 'GroupStatusBusy'
  204 = 'GroupStatusValid'
  973 = 'GroupStopping'
  680 = 'ID Detection Active'
  238 = 'ID Detection Error'
  526 = 'ID Detection Mode: %s'
  29 = 'ID Detection Valid'
  563 = 'In Target'
  211 = 'Info Act Pos Absolute'
  586 = 'Info Act Pos Modulo'
  21 = 'Info Mover Avoiding Collision'
  282 = 'Info Mover Coupled'
  398 = 'Info Mover Enabled'
  751 = 'Info Mover Error'
  907 = 'Info Mover Standstill'
  480 = 'Info nError ID'
  922 = 'Info Target Pos Absolute'
  16 = 'Info Target Pos Modulo'
  779 = 'Mask: %s'
  726 = 'McGroupState:      %s'
  974 = 'MOVER command'
  387 = 'Mover ID: %d'
  297 = 'Mover Position Assignement: %s'
  840 = 'MOVER result:  %s'
  53 = 'MOVER state:   %s'
  827 = 'nMask'
  145 = 'nMover: %d'
  825 = 'nMoverId'
  756 = 'nMoverSelected: %d'
  826 = 'nTargetStation'
  427 = 'Offset: %.3f'
  312 = 'Operation Mode: %s'
  320 = 'Queue: %d'
  828 = 'rOffset'
  642 = 'SelectBy:  %d'
  91 = 'Set Acceleration'
  399 = 'Set Delta'
  382 = 'Set Distance'
  757 = 'Set Gap'
  934 = 'Set Jerk'
  201 = 'Set Override'
  936 = 'Set Position'
  62 = 'Set Velocity'
  231 = 'State'
  567 = 'Target Station: %d'
  227 = 'XpuResult:   %s'
  96 = 'XpuState:    %s'
  884 = 'XTS Station'
  572 = 'XTS Transport Check:  %s'
  500 = 'XTS Transport Command'
  805 = 'XTS Transport Initialisation:  %s'
  395 = 'XTS Transport Result: %s'
  798 = 'XTS Transport State:  %s'
END_TEXTLIST

// ---- XTS_TRANSPORT/_Visualization/GROUP_VISU.TcVIS
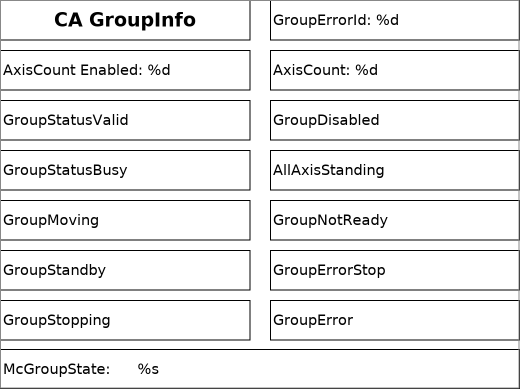
VISUALIZATION GROUP_VISU  // 520x389
VAR_IN_OUT
	stGroupInfo   : ST_GROUP_INFO;
  sGroupState   : string(60);
END_VAR
    Rectangle (0,100 250x40), "GroupStatusValid", colour toggle: stGroupInfo.GroupStatusValid
    Rectangle (0,150 250x40), "GroupStatusBusy", colour toggle: stGroupInfo.GroupStatusBusy
    Rectangle (0,200 250x40), "GroupMoving", colour toggle: stGroupInfo.GroupMoving
    Rectangle (270,250 250x40), "GroupErrorStop", colour toggle: stGroupInfo.GroupErrorStop
    Rectangle (270,200 250x40), "GroupNotReady", colour toggle: stGroupInfo.GroupNotReady
    Rectangle (0,250 250x40), "GroupStandby", colour toggle: stGroupInfo.GroupStandby
    Rectangle (0,300 250x40), "GroupStopping", colour toggle: stGroupInfo.GroupStopping
    Rectangle (270,100 250x40), "GroupDisabled", colour toggle: stGroupInfo.GroupDisabled
    Rectangle (270,150 250x40), "AllAxisStanding", colour toggle: stGroupInfo.AllAxesStanding
    Rectangle (270,300 250x40), "GroupError", colour toggle: stGroupInfo.GroupError
    Rectangle (270,0 250x40), "GroupErrorId: %d", text variable: stGroupInfo.GroupErrorId
    Rectangle (270,50 250x40), "AxisCount: %d", text variable: stGroupInfo.AxisCount
    Rectangle (0,349 520x40), "McGroupState: %s", text variable: sGroupState
    Rectangle (0,0 250x40), "CA GroupInfo"
    Rectangle (0,50 250x40), "AxisCount Enabled: %d", text variable: stGroupInfo.AxisCountEnabled
END_VISUALIZATION

// ---- XTS_TRANSPORT/_Visualization/textlists/TL_E_CTRL_MOVER.TcTLO
TEXTLIST TL_E_CTRL_MOVER
  0 = 'MOVER_NULL'
  1 = 'MOVER_ENABLE'
  2 = 'MOVER_DISABLE'
  4 = 'MOVER_MOVE_TO_POS_CA'
  5 = 'MOVER_SEND_TO_POS_CA'
  6 = 'MOVER_HALT'
  7 = 'MOVER_GEAR_IN'
  8 = 'MOVER_GEAR_IN_POS_CA'
  9 = 'MOVER_GEAR_OUT'
  10 = 'MOVER_RESET'
  3 = 'MOVER_MOVE_TO_POS'
   = ''
END_TEXTLIST

// ---- XTS_TRANSPORT/_Visualization/textlists/TL_E_CTRL_STATION.TcTLO
TEXTLIST TL_E_CTRL_STATION
  0 = 'STATION_CTRL_NULL'
  1 = 'STATION_INIT'
  10 = 'STATION_DISABLE'
  11 = 'STATION_ENABLE'
  20 = 'STATION_MOVER_ENTER'
  21 = 'STATION_MOVER_ENTER_RETRY'
  22 = 'STATION_MOVER_SEND'
  30 = 'STATION_PROCESS_START'
  31 = 'STATION_PROCESS_DONE'
  50 = 'STATION_MOVER_OUT'
  51 = 'STATION_MOVER_OUT_RETRY'
  60 = 'STATION_MOVER_GONE'
   = ''
END_TEXTLIST

// ---- XTS_TRANSPORT/_Visualization/textlists/TL_E_CTRL_TRANSPORT.TcTLO
TEXTLIST TL_E_CTRL_TRANSPORT
  0 = 'CMD_NULL'
  10 = 'CMD_INIT'
  11 = 'CMD_IDLE'
  20 = 'CMD_MOVER_ENABLE'
  21 = 'CMD_MOVER_DISABLE'
  22 = 'CMD_MOVER_HALT_CA'
  23 = 'CMD_MOVER_STOP'
  30 = 'CMD_GROUP_CLEAR'
  31 = 'CMD_GROUP_BUILD'
  32 = 'CMD_GROUP_ENABLE'
  33 = 'CMD_GROUP_STOP'
  40 = 'CMD_TRANSPORT_START'
  41 = 'CMD_TRANSPORT_RESTART'
   = ''
END_TEXTLIST

// ---- XTS_TRANSPORT/_Visualization/textlists/TL_E_CTRL_XPU.TcTLO
TEXTLIST TL_E_CTRL_XPU
  0 = 'XTS_CMD_NULL'
  10 = 'XTS_CMD_INIT'
  30 = 'XTS_IDLE'
   = ''
END_TEXTLIST

// ---- XTS_TRANSPORT/_Visualization/types/T_MOVER_SELECTOR.TcVIS
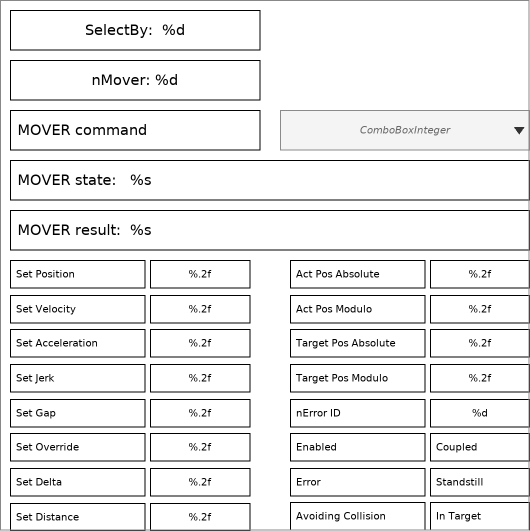
VISUALIZATION T_MOVER_SELECTOR  // 530x531
VAR_IN_OUT
	Control     : ST_MOVER_SELECTOR_CTRL;
  State       : ST_MOVER_SELECTOR_STATE;
  sState      : STRING;
  sResult     : STRING;
END_VAR
    Rectangle (10,60 250x40), "nMover: %d", text variable: Control.Mover
        OnMouseClick: write the text variable via VisuDialogs.Numpad, min 1, max MAX_MOVER, title 'Selected Mover'
    Rectangle (10,10 250x40), "SelectBy: %d", text variable: Control.Selector, text list: 'TL_E_MOVER_SELECTOR'
        p4168582468: "0 = SelectBy Index"
        OnMouseClick: write the text variable via VisuDialogs.Numpad, min 0, max 1, title 'SelectBy'
    Rectangle (10,160 520x40), "MOVER state: %s", text variable: sState
    Rectangle (10,110 250x40), "MOVER command"
    ComboBoxInteger (280,110 250x40), variable: Control.Control.Cmd, text list: 'TL_E_CTRL_MOVER'
    Rectangle (10,210 520x40), "MOVER result: %s", text variable: sResult
    Rectangle (10,260 135x28), "Set Position"
    Rectangle (10,295 135x28), "Set Velocity"
    Rectangle (10,329 135x28), "Set Acceleration"
    Rectangle (10,364 135x28), "Set Jerk"
    Rectangle (10,399 135x28), "Set Gap"
    Rectangle (10,433 135x28), "Set Override"
    Rectangle (10,468 135x28), "Set Delta"
    Rectangle (10,503 135x28), "Set Distance"
    Rectangle (150,260 100x28), "%.2f", text variable: Control.Data.rPos
        OnMouseClick: write the text variable via Default
    Rectangle (150,295 100x28), "%.2f", text variable: Control.Data.rVelo
        OnMouseClick: write the text variable via Default
    Rectangle (150,329 100x28), "%.2f", text variable: Control.Data.rAcc
        OnMouseClick: write the text variable via Default
    Rectangle (150,364 100x28), "%.2f", text variable: Control.Data.rJerk
        OnMouseClick: write the text variable via Default
    Rectangle (150,399 100x28), "%.2f", text variable: Control.Data.rGap
        OnMouseClick: write the text variable via Default
    Rectangle (150,433 100x28), "%.2f", text variable: Control.Data.rOverride
        OnMouseClick: write the text variable via Default
    Rectangle (150,468 100x28), "%.2f", text variable: Control.Data.rDelta
        OnMouseClick: write the text variable via Default
    Rectangle (150,503 100x28), "%.2f", text variable: Control.Data.rDistance
        OnMouseClick: write the text variable via Default
    Rectangle (290,260 135x28), "Act Pos Absolute"
    Rectangle (290,295 135x28), "Act Pos Modulo"
    Rectangle (290,329 135x28), "Target Pos Absolute"
    Rectangle (290,364 135x28), "Target Pos Modulo"
    Rectangle (290,399 135x28), "nError ID"
    Rectangle (430,260 100x28), "%.2f", text variable: State.Info.rAbsActPos
    Rectangle (430,295 100x28), "%.2f", text variable: State.Info.rModuloActPos
    Rectangle (430,329 100x28), "%.2f", text variable: State.Info.rAbsTargetPos
    Rectangle (430,364 100x28), "%.2f", text variable: State.Info.rModuloTargetPos
    Rectangle (430,399 100x28), "%d", text variable: State.Info.nErrorId
    Rectangle (290,433 135x28), "Enabled", colour toggle: State.Info.bMoverEnabled
    Rectangle (290,468 135x28), "Error", colour toggle: State.Info.bMoverError
    Rectangle (430,433 100x28), "Coupled", colour toggle: State.Info.bMoverCoupled
    Rectangle (430,468 100x28), "Standstill", colour toggle: State.Info.bMoverStandstill
    Rectangle (290,502 135x28), "Avoiding Collision", colour toggle: State.Info.bMoverAvoidingCollision
    Rectangle (430,502 100x28), "In Target", colour toggle: State.Info.bMoverInTarget
END_VISUALIZATION

// ---- XTS_TRANSPORT/_Visualization/XPU_VISU.TcVIS
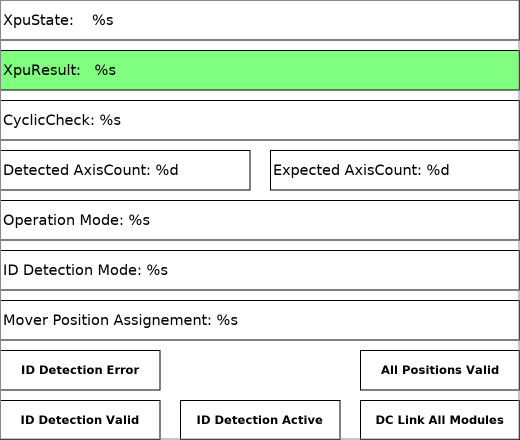
VISUALIZATION XPU_VISU  // 520x440
VAR_IN_OUT
	stXpuState    : ST_XPU_STATE;
  stXpuInfo     : ST_XPU_INFO;
  stXpuStrings  : ST_XPU_STRINGS;
END_VAR
    Rectangle (0,100 520x40), "CyclicCheck: %s", text variable: stXpuStrings.sXpuCyclicCheck
    Rectangle (0,0 520x40), "XpuState: %s", text variable: stXpuStrings.sXpuState
    Rectangle (0,50 520x40), "XpuResult: %s", text variable: stXpuStrings.sXpuResult, colour toggle: (MAIN.eXpuResult = E_PROGRESS.PROGRESS_ERROR)
    Rectangle (360,350 160x40), "All Positions Valid", colour toggle: stXpuInfo.AllPositionsValid
    Rectangle (0,350 160x40), "ID Detection Error", colour toggle: stXpuInfo.IdDetectionError
    Rectangle (0,400 160x40), "ID Detection Valid", colour toggle: stXpuInfo.IdDetectionValid
    Rectangle (180,400 160x40), "ID Detection Active", colour toggle: stXpuInfo.IdDetectionActive
    Rectangle (0,200 520x40), "Operation Mode: %s", text variable: stXpuStrings.sXpuOpMode
    Rectangle (0,250 520x40), "ID Detection Mode: %s", text variable: stXpuStrings.sXpuMoverId_DetectionMode
    Rectangle (0,300 520x40), "Mover Position Assignement: %s", text variable: stXpuStrings.sXpuMoverPosAssignement
    Rectangle (270,150 250x40), "Expected AxisCount: %d", text variable: stXpuInfo.nExpectedAxisCount
    Rectangle (0,150 250x40), "Detected AxisCount: %d", text variable: stXpuInfo.nDetectedAxisCount
    Rectangle (360,400 160x40), "DC Link All Modules", colour toggle: stXpuState.DcLink
END_VISUALIZATION

// ---- _MSG/types/TL_E_MESSAGETYPE.TcTLO
TEXTLIST TL_E_MESSAGETYPE
  0 = 'eMessageEmpty'
  1 = 'eMessageError'
  2 = 'eMessageWarning'
  3 = 'eMessageInfo'
  4 = 'eMessageVerbose'
   = ''
END_TEXTLIST
